(* IEC 61131-3 sources: 2026_Projet_YGO_ExcavatriceDragage/CODE_BACKUP/CODE_20260904_AvantWeekendBackup_v0.6.34/G_CYCLE (part 2) *)

(* ---- FB_CycleSemiAuto.st ---- *)
(* =======================================================================
   ⚙️ FB_CycleSemiAuto — Séquenceur du cycle automatique (Grafcet de dragage)
   ───────────────────────────────────────────────────────────────
   🎯 Rôle : Automate de cycle automatique de dragage (X0 à X13 + AX_STAB)
   🔒 Sécurité : Gating par mode et homme-mort, repli AX_STAB sur défaut
   🔌 Interface : Demandes de mouvements (treuils, translation, benne)
   📄 Doc métier : DOC/AF/AF_Partie-04_Mode_SemiAuto_Sequenceur_v2.3.md
   ======================================================================= *)

FUNCTION_BLOCK PUBLIC FB_CycleSemiAuto
VAR_INPUT
    // === COMMANDES & AUTORISATIONS ===
    Enable                  : BOOL;         // --> [CMD] Activation generale du sequenceur
    Reset                   : BOOL;         // --> [CMD] Acquittement defaut (front)
    PowerContactorEngaged   : BOOL;         // --> [SAFE] Chaine de securite OK
    EncoderFaultPresent     : BOOL;         // --> [SAFE] Defaut codeur agrege (cycle non autorise)
    Mode                    : E_Mode;       // --> [CMD] Mode arbitre (SEMI_AUTO pour instance cycle)
    JoystickDeflected       : BOOL;         // --> [CMD] Manche deflecte (non centre)
    DeadmanArmed            : BOOL;         // --> [CMD] Appui homme-mort (fenetre 3 s)
    HeartbeatIhmOk          : BOOL;         // --> [SAFE] IHM<->PLC valide

    // === COMMANDES OPERATEUR ===
    StartCycle              : BOOL;         // --> [CMD] Demande lancement / reprise (IHM)
    AbortCycle              : BOOL;         // --> [CMD] Demande abandon (IHM)

    // === CIBLES ET CONFIGURATION ===
    SelTarget               : INT;          // --> [CFG] RESERVE (C3.1 : le cycle part toujours de P1, plus de selection de cible). Cable, non consomme.
    SetDepthM               : REAL;         // --> [CFG] Profondeur de consigne (negative)
    SetOffsetM              : REAL;         // --> [CFG] Ecart de fermeture benne cible

    // === FEEDBACKS CAPTEURS & MATERIEL ===
    KoboldContactFond       : BOOL;         // --> [HW] Retour dedie Kobold : TRUE = contact fond (front descendant DI)
    KoboldImmersed          : BOOL;         // --> [HW] Etat brut DI Kobold : TRUE = sonde dans l'eau (fronts AX6/AX7)
    KoboldContactorFeedback : BOOL;         // --> [HW] Retour contacteur Kobold enclenche (verif init AX5)
    LimitLegalReached       : BOOL;         // --> [SAFE] Limite legale atteinte (descente interdite)
    LimitLegalDepthM        : REAL;         // --> [CFG] Profondeur legale minimale autorisee
    WinchSyncError          : BOOL;         // --> [SAFE] Desynchronisme bloquant M1/M2
    WinchSyncDeltaM         : REAL;         // --> [HW] Ecart codeurs M1/M2 pour diagnostic
    M1_CablePosM            : REAL;         // --> [HW] Position cable treuil M1 (recalee)
    M2_CablePosM            : REAL;         // --> [HW] Position cable treuil M2 (recalee)
    M1_MeasuredSpeedMps     : REAL;         // --> [HW] Vitesse lineaire mesuree M1 (m/s)
    M2_MeasuredSpeedMps     : REAL;         // --> [HW] Vitesse lineaire mesuree M2 (m/s)
    SpeedMismatchThresholdMps : REAL;       // --> [CFG] Seuil ecart vitesse ; 0 = controle desactive
    SpeedMismatchTimeout    : TIME;         // --> [CFG] Duree de confirmation ; 0 = controle desactive
    CableLimitM1AscentM     : REAL;         // --> [CFG] Limite haute d'exploitation M1

    // === FEEDBACKS TRANSLATION M3 ===
    Translation_At_P1           : BOOL;     // --> [HW] Capteur position P1 (arret travail)
    Translation_At_Tremie       : BOOL;     // --> [HW] Capteur fin de course tremie
    Translation_At_Maintenance : BOOL;     // --> [HW] Capteur fin de course maintenance
    Translation_Busy            : BOOL;     // --> [HW] Mouvement translation en cours
    Translation_Done            : BOOL;     // --> [HW] Cible translation atteinte

    // === FEEDBACKS BENNE ===
    Benne_Busy              : BOOL;         // --> [HW] Mouvement machoires benne en cours
    Benne_Done              : BOOL;         // --> [HW] Mouvement ouverture/fermeture termine
    Benne_IsOpen            : BOOL;         // --> [HW] Benne mecaniquement ouverte memorisee
    Benne_IsClosed          : BOOL;         // --> [HW] Benne mecaniquement fermee memorisee
    Benne_IsRoughlyClosed   : BOOL;         // --> [HW] Benne a peu pres fermee (tolerance matiere)

    // === REFERENCEMENT CODEURS ===
    HomedM1                 : BOOL;         // --> [HW] Codeur M1 reference
    HomedM2                 : BOOL;         // --> [HW] Codeur M2 reference
    TopPositionSensor       : BOOL;         // --> [HW] Capteur position haute (referencement)
    HomingRequest           : BOOL;         // --> [CMD] Demande de referencement (front)
    InitPositionOk          : BOOL;         // --> [HW] Posture de depart OK (treuils/M3 dans la plage, calcul PRG_03) - condition AX1_INIT
    WinchesAtTopWindow      : BOOL;         // --> [HW] Treuils M1 ET M2 dans la fenetre FDC logiciel haut (calcul PRG_03) - surveille en AX2

    // === CONFIG & COMMANDES CYCLE (IHM) ===
    CfgDrainTime           : TIME;         // --> [CFG] Duree d'egouttage AX13 configurable IHM (<= 0 -> defaut interne)
    SkipDrainRequest       : BOOL;         // --> [CMD] Bouton IHM : passer l'etape d'egouttage AX13 (front)
    RepositionRequest      : BOOL;         // --> [CMD] Option IHM (maintenue) : repositionnement couple M1+M2 pendant le vidage tremie (AX15B <-> AX15C)

    // === CONFIG DIVING / EXTRACTION (GEL 2026-09-03) ===
    DiveStartMinM          : REAL;         // --> [CFG] Altimetrie de lancement Kobold (AT4 : AX4 -> AX5), reglable IHM (~3..5 m ; <= 0 -> defaut interne)
    CfgRaiseOffBottomM     : REAL;         // --> [CFG] Decollement du fond en AX8 : RaiseTargetM = TouchPositionM + ce champ (reglable IHM ; <= 0 -> 0,5 m)
    CfgCtrlAscentMaxStep   : INT;          // --> [CFG] Palier max montee controle AX11, borne [1..2] (defaut 1)
    M1_SpeedStepApplied    : INT;          // --> [HW] Palier vitesse effectivement applique M1 (0 = inconnu ; garde palier <> 4 en diving)
    M2_SpeedStepApplied    : INT;          // --> [HW] Palier vitesse effectivement applique M2 (0 = inconnu)
END_VAR
VAR_OUTPUT
    // === ETATS IEC & DEFECTUOSITES ===
    Ready                   : BOOL;         // <-- [STAT] Sequenceur disponible
    Fault                   : ST_Fault;     // <-- [SAFE] Socle defaut transverse (live + latche)
    Lifecycle               : ST_Lifecycle; // <-- [STAT] Cycle de vie (Busy, Done, Waiting)
    SpeedMismatchMps        : REAL;         // <-- [DIAG] Ecart absolu vitesse M1/M2 (m/s)
    SpeedMismatchActive     : BOOL;         // <-- [DIAG] Seuil vitesse depasse sur cycle courant
    SpeedMismatchConfirmed  : BOOL;         // <-- [DIAG] Ecart vitesse confirme pendant timeout
    BottomTouched           : BOOL;         // <-- [STAT] Fond touche (latch AX8, efface a AX0 / AX_STAB / Reset) - variable d'info GEL AX8

    // === ORDRES ACTIONNEURS (COMMANDES STRUCTUREES) ===
    // Types de contrat inter-PRG uniques (ST_Program*Request) : FB_CycleSemiAuto produit
    // directement les demandes consommées par PRG_04/05/07 — plus de DUT
    // ST_fbCycle_*CmdDemand redondants ni de re-mapping champ-à-champ (NC-090).
    WinchM1Cmd              : ST_ProgramWinchRequest;        // <-- [ACT] Demande treuil M1
    WinchM2Cmd              : ST_ProgramWinchRequest;        // <-- [ACT] Demande treuil M2
    TranslationCmd          : ST_ProgramTranslationRequest;  // <-- [ACT] Demande translation M3
    BucketCmd               : ST_ProgramBucketRequest;       // <-- [ACT] Demande benne

    // === METADONNEES & SYNOPTIQUE ===
    CycleStep               : E_AutoCycleStep;          // <-- [STAT] Etape active du Grafcet
    CycleStateStr           : STRING(80);           // <-- [STAT] Libelle en clair de l'etape
    CycleStepAtError        : E_AutoCycleStep;          // <-- [DIAG] Etape specifique au moment du defaut
    OperatorActionId        : WORD;                 // <-- [DIAG] ID action operateur requise
    OperatorAction          : STRING(120);          // <-- [DIAG] Message explicatif pour l'IHM
    ExpectedAxis            : E_OperatorAxis;       // <-- [STAT] Organe joystick/bouton attendu
    ExpectedDirection       : INT;                  // <-- [STAT] Sens attendu (-1, 0, +1)
    WaitingForOperator      : BOOL;                 // <-- [STAT] En attente d'une action operateur
    WaitingForProcess       : BOOL;                 // <-- [STAT] En attente d'une condition procede
    RequestActive           : BOOL;                 // <-- [STAT] Demande de mouvement active
    CurrentCycleElapsed     : TIME;                 // <-- [DIAG] Duree ecoulee du cycle en cours (chronometre sur Lifecycle.Busy)
    LastCycleDuration       : TIME;                 // <-- [DIAG] Duree du dernier cycle acheve (figee a X13, persiste au cycle suivant)
END_VAR
VAR_IN_OUT
    // === STRUCTURES PARTAGEES & COMPTEURS ===
    SampleCount             : INT;          // <-> [BUS] Compteur de prelevements (RETAIN)
END_VAR
VAR
    // === DETECTEURS DE FRONTS ===
    ResetEdge               : R_TRIG;       // . [LOC] Detecteur front montant Reset
    StartEdge               : R_TRIG;       // . [LOC] Detecteur front montant StartCycle
    DeadmanArmedEdge        : R_TRIG;       // . [LOC] Detecteur front montant DeadmanArmed (demarrage joystick)
    AbortEdge               : R_TRIG;       // . [LOC] Detecteur front montant AbortCycle
    ErrorEdge               : R_TRIG;       // . [LOC] Detecteur front montant Error
    JoyDeflectedEdge        : R_TRIG;       // . [LOC] Front montant JoystickDeflected (relance AX18 sur geste franc, pas maintien)

    // === GATE CONTINU HOMME-MORT ===
    CycleMotionPermit       : BOOL; // . [LOC] Permis de mouvement cycle = JoystickDeflected AND DeadmanArmed (manche deflechi + homme-mort arme) ; gate commun a toutes les commandes d'actionneur du sequenceur. Le sens du mouvement reste porte par ReqAscent/ReqDescend de chaque etape.

    // === COMPTEUR PRELEVEMENTS (garde de front) ===
    SampleCountDone         : BOOL := FALSE; // . [LOC] F2: front de comptage SampleCount (1 seul increment par cycle)

    // === ETATS INTERNES ===
    State                   : E_AutoCycleStep := E_AutoCycleStep.AX0_REPOS; // . [LOC] Etape courante machine d'etat
    SavedState              : E_AutoCycleStep := E_AutoCycleStep.AX0_REPOS; // . [LOC] Etape memorisee
    PausedState             : E_AutoCycleStep := E_AutoCycleStep.AX0_REPOS; // . [LOC] Etape en pause lors de la bascule hors auto
    WaitingResume           : BOOL := FALSE;                             // . [LOC] En attente de validation consciente pour reprendre

    // === MEMORISATIONS & REGISTRES INTERNES ===
    TouchPositionM          : REAL;         // . [LOC] Position M1 memorisee lors du contact fond
    RaiseTargetM            : REAL;         // . [LOC] Profondeur de remontee memorisee
    SelectedWorkTarget      : INT;          // . [LOC] Cible de travail (fige a 3=P1 depuis C3.1) - conserve pour diag/futur
    InitConditionsOk        : BOOL;         // . [LOC] AX1_INIT : toutes les conditions initiales sont remplies
    StepMaxPrevState        : E_AutoCycleStep;  // . [LOC] Etape du scan precedent (rearmement StepMaxTimer au changement d'etape)

    // === FRONTS / TEMPO DIVING ===
    KoboldRiseEdge          : R_TRIG;       // . [LOC] Front DI Kobold 0->1 (entree dans l'eau, AX6)
    KoboldFallEdge          : F_TRIG;       // . [LOC] Front DI Kobold 1->0 (fond, AX7)
    KoboldInitTimer         : TON;          // . [LOC] Fenetre de verif retour contacteur Kobold en AX5
    RetryJoyReleaseTimer    : TON;          // . [LOC] Anti-rebond relache joystick pendant diving (>= 200 ms avant reprise)
    PalierNot4Timer         : TON;          // . [LOC] Confirmation palier bloque < 4 en plongee (tolere la rampe 1->4)
    DivingRetryTrig         : BOOL;         // . [LOC] Synthese GT-dive-retry (erreur Kobold / joystick relache / palier < 4 confirme en AX5..AX7)
    CtrlAscentMaxStepEff    : INT;          // . [LOC] CfgCtrlAscentMaxStep borne [1..2]
    RaiseOffBottomEff       : REAL;         // . [LOC] CfgRaiseOffBottomM borne (>0, defaut 0,5 m)
    DiveStartMinEff         : REAL;         // . [LOC] DiveStartMinM borne (defaut interne si <= 0)

    // === TEMPORISATEURS INTERNES ===
    DrainingTimer           : TON;          // . [LOC] Temporisateur de vidage (egouttage), PT = DrainTimeEff
    CycleRunTimer           : TON;          // . [LOC] Chronometre du cycle en cours (IN = Lifecycle.Busy) ; .ET = duree
    SkipDrainEdge           : R_TRIG;       // . [LOC] Front bouton IHM "passer egouttage"
    DrainTimeEff            : TIME;         // . [LOC] Duree d'egouttage effective (CfgDrainTime bornee au defaut interne)
    StabilizationTimer      : TON;          // . [LOC] Temporisation maximale de remontee lente
    SpeedMismatchTimer      : TON;          // . [LOC] Confirmation temporelle ecart de vitesse
    StepMaxTimer            : TON;          // . [LOC] Tempo max d'etape

    // === CONSTANTES & CONFIGURATIONS INTERNES ===
    CtrlAscentDistM         : REAL := 2.0;      // . [LOC] Distance de remontee lente de controle
    CtrlAscentToleranceM    : REAL := 0.25;     // . [LOC] Ecart maximal admis entre codeurs
    CtrlAscentTimeout       : TIME := T#30s;    // . [LOC] Temps max pour zone de stabilisation
    DrainingTime            : TIME := T#5s;     // . [LOC] Temps d'egouttage par defaut
    StepMaxTimeout          : TIME := T#60s;    // . [LOC] Tempo max d'etape

    // === SOCLE DEFAUT TRANSVERSE ===
    instFault               : FB_FaultCore;                  // * [INST] Socle defaut transverse
    instCauses              : ARRAY[0..15] OF ST_FaultCause; // . [LOC] Table des causes de defaut
END_VAR
VAR CONSTANT
    // Paliers de vitesse treuil par etape (StepTgt des demandes WinchMxCmd, 1..5 ; 0 = arret).
    CST_StepSlow   : INT := 1;   // Palier lent : retente AX9, controle AX11, repositionnement AX15C
    CST_StepDive   : INT := 4;   // Palier plongee Kobold AX4..AX7 : palier 4 MINI ET MAXI impose, palier 5 interdit (GEL Q9)
    CST_StepLoaded : INT := 4;   // Palier montee en charge AX12 (bridage strict <= 4, jamais palier 5)
    CST_KoboldInitTimeout : TIME := T#3s;   // Fenetre max de confirmation retour contacteur Kobold en AX5
    CST_RaiseOffBottomDefaultM : REAL := 0.5;   // Decollement du fond par defaut (AX8) si CfgRaiseOffBottomM <= 0
    // Backstop anti-telescopage : ecart de position M1/M2 max tolere pendant les phases
    // reellement couplees hors X7 (qui a deja son propre controle a 0,25 m). Aligne sur
    // CfgSyncCriticalToleranceM = 0,50 m (AF-04 §5). FB_SyncDeviation (PRG_04) reste la
    // surveillance primaire ; ceci est un garde-fou local au sequenceur.
    CST_CoupledPosBacklashM : REAL := 0.5;
END_VAR

// === IMPLEMENTATION ===

{region "§1 Causes & Socle Défaut"}
// 🔑 1. FRONTS ET CAUSES
ResetEdge(CLK := Reset);
StartEdge(CLK := StartCycle);
DeadmanArmedEdge(CLK := DeadmanArmed);
AbortEdge(CLK := AbortCycle);
SkipDrainEdge(CLK := SkipDrainRequest);
KoboldRiseEdge(CLK := KoboldImmersed);
KoboldFallEdge(CLK := KoboldImmersed);
JoyDeflectedEdge(CLK := JoystickDeflected);

// Config diving/extraction bornee (repli defaut interne si non reglee / valeur implausible).
// DiveStartMinM = altimetrie de lancement Kobold dans le referentiel M1_CablePosM
// (positif, ~7,5 m au FDC haut, decroissant a la descente). Plage plausible 0,5..8,0 m ;
// hors plage -> repli 4,0 m.
IF (DiveStartMinM >= 0.5) AND (DiveStartMinM <= 8.0) THEN
    DiveStartMinEff := DiveStartMinM;
ELSE
    DiveStartMinEff := 4.0;
END_IF;
RaiseOffBottomEff := SEL(CfgRaiseOffBottomM > 0.0, CST_RaiseOffBottomDefaultM, CfgRaiseOffBottomM);
CtrlAscentMaxStepEff := LIMIT(1, CfgCtrlAscentMaxStep, 2);

// ⏱️ Chronomètre du cycle : compte tant que le séquenceur est actif (Lifecycle.Busy).
// .ET = durée écoulée du cycle en cours ; figée dans LastCycleDuration à l'achèvement (X13).
CycleRunTimer(IN := Lifecycle.Busy, PT := T#12h);
CurrentCycleElapsed := CycleRunTimer.ET;

// Durée d'égouttage effective : config IHM si valide, sinon défaut interne.
DrainTimeEff := SEL(CfgDrainTime <= T#0s, CfgDrainTime, DrainingTime);

// ⏱️ Surveillance indépendante de la remontée lente de controle
// AX11_CTRL_ASCENT -> AX12_LOADED_ASCENT : TON de stabilisation palier lent.
StabilizationTimer(IN := (State = E_AutoCycleStep.AX11_CTRL_ASCENT), PT := CtrlAscentTimeout);

// ⏱️ AX5_KOBOLD_INIT : fenetre de confirmation du retour contacteur Kobold.
KoboldInitTimer(IN := (State = E_AutoCycleStep.AX5_KOBOLD_INIT), PT := CST_KoboldInitTimeout);

// 📏 Comparaison vitesse réelle M1/M2
SpeedMismatchMps := ABS(M1_MeasuredSpeedMps - M2_MeasuredSpeedMps);
SpeedMismatchActive := (State = E_AutoCycleStep.AX11_CTRL_ASCENT)
                       AND JoystickDeflected
                       AND (SpeedMismatchThresholdMps > 0.0)
                       AND (SpeedMismatchTimeout > T#0ms)
                       AND (SpeedMismatchMps > SpeedMismatchThresholdMps);
// AX11_CTRL_ASCENT -> AX_STAB : TON confirmation écart vitesse.
SpeedMismatchTimer(IN := SpeedMismatchActive, PT := SpeedMismatchTimeout);
SpeedMismatchConfirmed := SpeedMismatchTimer.Q;

// Tempo max d'étape (R5) — backstop durée d'état, lancé SEULEMENT si pilotage joystick actif.
// Xi -> AX_STAB sur dépassement. Réarmé à CHAQUE changement d'étape (IN=FALSE 1 scan) :
// chaque étape dispose de sa propre fenêtre StepMaxTimeout, la tempo n'est PAS cumulative
// sur l'ensemble du cycle (un cycle réel long ne tombe plus en AX_STAB intempestif).
StepMaxTimer(IN := (State = StepMaxPrevState)
                  AND JoystickDeflected
                  AND (State <> E_AutoCycleStep.AX0_REPOS)
                  AND (State <> E_AutoCycleStep.AX18_DONE_SYNC)
                  AND (State <> E_AutoCycleStep.AX_STAB)
                  AND (State <> E_AutoCycleStep.AX_DIVING_RETRY),
             PT := StepMaxTimeout);
StepMaxPrevState := State;

// Egouttage AX13 : TON gaté sur l'étape (remis à 0 hors AX13). Remplace l'ancien IN:=TRUE câblé
// qui pouvait laisser Q déjà vrai à l'entrée en AX13 (temps d'égouttage non respecté).
DrainingTimer(IN := (State = E_AutoCycleStep.AX13_DRAIN_PAUSE), PT := DrainTimeEff);

// GT-dive-retry (GEL Q11) : en AX5/AX6/AX7, erreur sequence Kobold (retour contacteur
// absent apres CST_KoboldInitTimeout) OU joystick relache (>= 200 ms, anti-rebond) OU
// palier applique <> 4 sur M1 ou M2 (feedback si cable) -> reprise AX_DIVING_RETRY
// (PAS un defaut latche).
RetryJoyReleaseTimer(IN := ((State = E_AutoCycleStep.AX5_KOBOLD_INIT)
                             OR (State = E_AutoCycleStep.AX6_SEARCH_IMMERSION)
                             OR (State = E_AutoCycleStep.AX7_SEARCH_BOTTOM))
                            AND NOT JoystickDeflected,
                     PT := T#200ms);
// Palier bloque SOUS 4 pendant la plongee : on TOLERE la rampe 1->4 (tempo contacteurs,
// GEL AX4) ; seul un blocage confirme > 4 s en AX5..AX7 declenche la reprise. Palier 5
// (> 4) est traite instantanement par la cause de defaut 8 (latche), pas ici.
PalierNot4Timer(IN := ((State = E_AutoCycleStep.AX5_KOBOLD_INIT)
                        OR (State = E_AutoCycleStep.AX6_SEARCH_IMMERSION)
                        OR (State = E_AutoCycleStep.AX7_SEARCH_BOTTOM))
                       AND JoystickDeflected
                       AND ( ((M1_SpeedStepApplied > 0) AND (M1_SpeedStepApplied < CST_StepDive))
                          OR ((M2_SpeedStepApplied > 0) AND (M2_SpeedStepApplied < CST_StepDive)) ),
                PT := T#5s);
DivingRetryTrig := ((State = E_AutoCycleStep.AX5_KOBOLD_INIT)
                     OR (State = E_AutoCycleStep.AX6_SEARCH_IMMERSION)
                     OR (State = E_AutoCycleStep.AX7_SEARCH_BOTTOM))
                   AND ( (KoboldInitTimer.Q AND NOT KoboldContactorFeedback)
                         OR RetryJoyReleaseTimer.Q
                         OR PalierNot4Timer.Q );

// Table des causes de défaut
instCauses[0].Active   := LimitLegalReached
                          AND ((State = E_AutoCycleStep.AX4_DESCEND_DIVING)
                            OR (State = E_AutoCycleStep.AX5_KOBOLD_INIT)
                            OR (State = E_AutoCycleStep.AX6_SEARCH_IMMERSION)
                            OR (State = E_AutoCycleStep.AX7_SEARCH_BOTTOM));
instCauses[0].Latching := TRUE;
instCauses[0].Texte    := 'Limite legale de profondeur atteinte pendant descente';

instCauses[1].Active   := WinchSyncError AND (State <> E_AutoCycleStep.AX0_REPOS) AND (State <> E_AutoCycleStep.AX_STAB);
instCauses[1].Latching := TRUE;
instCauses[1].Texte    := 'Desynchronisme treuils M1/M2 bloquant';

instCauses[2].Active   := SpeedMismatchConfirmed AND (State <> E_AutoCycleStep.AX0_REPOS) AND (State <> E_AutoCycleStep.AX_STAB);
instCauses[2].Latching := TRUE;
instCauses[2].Texte    := 'Ecart de vitesse M1/M2 confirme en montee';

instCauses[3].Active   := NOT HeartbeatIhmOk AND (State <> E_AutoCycleStep.AX0_REPOS) AND (State <> E_AutoCycleStep.AX_STAB);
instCauses[3].Latching := TRUE;
instCauses[3].Texte    := 'Perte communication IHM pendant cycle';

instCauses[4].Active   := StepMaxTimer.Q AND (State <> E_AutoCycleStep.AX_STAB);
instCauses[4].Latching := TRUE;
instCauses[4].Texte    := 'Depassement tempo maximale d etape (blocage mouvement)';

instCauses[5].Active   := (StabilizationTimer.Q OR (ABS(M1_CablePosM - M2_CablePosM) > CtrlAscentToleranceM))
                          AND (State = E_AutoCycleStep.AX11_CTRL_ASCENT);
instCauses[5].Latching := TRUE;
instCauses[5].Texte    := 'Defaut de stabilisation / tolerance ecart codeurs en remontee controle';

// Backstop anti-telescopage : ecart de position M1/M2 excessif pendant une phase
// reellement couplee. AX11 a deja son propre controle (instCauses[5]). Seuil grossier
// (0,50 m) : filet local si FB_SyncDeviation (PRG_04) ne coupe pas.
instCauses[6].Active   := (ABS(M1_CablePosM - M2_CablePosM) > CST_CoupledPosBacklashM)
                          AND JoystickDeflected
                          AND ((State = E_AutoCycleStep.AX4_DESCEND_DIVING)
                            OR (State = E_AutoCycleStep.AX5_KOBOLD_INIT)
                            OR (State = E_AutoCycleStep.AX6_SEARCH_IMMERSION)
                            OR (State = E_AutoCycleStep.AX7_SEARCH_BOTTOM)
                            OR (State = E_AutoCycleStep.AX9_RAISE_OFF_BOTTOM)
                            OR (State = E_AutoCycleStep.AX12_LOADED_ASCENT)
                            OR (State = E_AutoCycleStep.AX15C_DUMP_REPOSITION));
instCauses[6].Latching := TRUE;
instCauses[6].Texte    := 'Ecart de position M1/M2 excessif en phase couplee (anti-telescopage)';

// AX2 : pendant la translation vers P1 les treuils M1/M2 doivent RESTER au FDC
// logiciel haut (WinchesAtTopWindow, calcul PRG_03). S'ils quittent la fenetre
// -> defaut latche, sortie cycle (GEL SEMI_AUTO cause 7 / Q10).
instCauses[7].Active   := NOT WinchesAtTopWindow AND (State = E_AutoCycleStep.AX2_TRANSLATE_P1);
instCauses[7].Latching := TRUE;
instCauses[7].Texte    := 'Treuils M1/M2 hors FDC haut pendant la translation vers P1';

// GEL cause 8 : palier vitesse > 4 (palier 5) applique pendant la plongee. Le FB commande
// toujours CST_StepDive = 4 ; un palier 5 en retour feedback = anomalie aval -> defaut latche.
// (Un palier < 4 en retour est traite en reprise par GT-dive-retry, pas ici.)
instCauses[8].Active   := (((M1_SpeedStepApplied > CST_StepDive) OR (M2_SpeedStepApplied > CST_StepDive)))
                          AND ((State = E_AutoCycleStep.AX4_DESCEND_DIVING)
                            OR (State = E_AutoCycleStep.AX5_KOBOLD_INIT)
                            OR (State = E_AutoCycleStep.AX6_SEARCH_IMMERSION)
                            OR (State = E_AutoCycleStep.AX7_SEARCH_BOTTOM));
instCauses[8].Latching := TRUE;
instCauses[8].Texte    := 'Palier vitesse > 4 (palier 5) pendant la plongee - interdit';

// Appel du socle de défaut
instFault(Enable := Enable, Reset := Reset, Causes := instCauses);
Fault := instFault.Fault;
ErrorEdge(CLK := Fault.Error);
{endregion}

{region "§2 Gate securite & Bascule Mode"}
// 🛑 2. GATES DE SÉCURITÉ ET NEUTRALISATION
// Le mode SEMI_AUTO peut être sélectionné sous AU/défaut (FB_Modes), mais le cycle
// ne tourne JAMAIS sans puissance (PowerContactorEngaged) ni avec un codeur défaillant
// (EncoderFaultPresent) — les données de position invalides rendraient le Grafcet erroné.
IF NOT Enable OR NOT PowerContactorEngaged OR EncoderFaultPresent THEN
    WinchM1Cmd.RunRequest     := FALSE;
    WinchM1Cmd.ReqAscent      := FALSE;
    WinchM1Cmd.ReqDescend     := FALSE;
    WinchM1Cmd.StepTgt        := 0;

    WinchM2Cmd.RunRequest     := FALSE;
    WinchM2Cmd.ReqAscent      := FALSE;
    WinchM2Cmd.ReqDescend     := FALSE;
    WinchM2Cmd.StepTgt        := 0;

    TranslationCmd.ReqStart   := FALSE;
    TranslationCmd.PositionTgt  := 0;

    BucketCmd.ReqOpen         := FALSE;
    BucketCmd.ReqClose        := FALSE;
    BucketCmd.ReqKoboldMeasureEnable := FALSE;

    // Si on quitte le semi-auto alors qu'un cycle était en cours, on mémorise l'étape pour la pause
    IF (State <> E_AutoCycleStep.AX0_REPOS) AND (State <> E_AutoCycleStep.AX18_DONE_SYNC) AND (State <> E_AutoCycleStep.AX_STAB) THEN
        PausedState := State;
        WaitingResume := TRUE;
    END_IF;

    CycleStep            := State;
    CycleStateStr        := 'Cycle desactive : securite/codeur/mode';
    Ready                := FALSE;
    Lifecycle.Busy       := FALSE;
    Lifecycle.Done       := FALSE;
    SpeedMismatchTimer(IN := FALSE, PT := SpeedMismatchTimeout);
    SpeedMismatchMps := 0.0;
    SpeedMismatchActive := FALSE;
    SpeedMismatchConfirmed := FALSE;
    OperatorActionId := 0;
    IF EncoderFaultPresent THEN
        OperatorAction := 'Cycle non autorise : defaut codeur present. Reinitialiser le defaut codeur.';
    ELSE
        OperatorAction := 'Passer en mode Semi-Auto et engager la securite pour activer le cycle.';
    END_IF;
    ExpectedAxis := E_OperatorAxis.NONE;
    ExpectedDirection := 0;
    WaitingForOperator := FALSE;
    WaitingForProcess := FALSE;
    RequestActive := FALSE;
    RETURN;
END_IF;

Ready := Enable AND NOT Fault.Latched;

// 🛡️ Gate continu homme-mort : le mouvement n'est autorisé que si le manche est
// défléchi (JoystickDeflected) ET l'homme-mort est armé (DeadmanArmed). Chaque
// commande de mouvement est gatée par ce permis à chaque scan (pas seulement au
// démarrage). Le séquenceur (transitions X0→X13) reste piloté par JoystickDeflected.
CycleMotionPermit := JoystickDeflected AND DeadmanArmed;

// Au retour en Semi-Auto, si une étape était en cours, on exige une reprise consciente
IF WaitingResume THEN
    // 🔒 Sécurité anti-redémarrage automatique (AF-04 §4.1) : le cycle ne reprend
    // PAS sur manche + homme-mort seuls. Il reste en attente d'un geste conscient
    // (StartCycle) avant de restaurer l'étape mémorisée.
    IF StartEdge.Q THEN
        State := PausedState;   // reprise consciente : restaure l'étape mémorisée
        WaitingResume := FALSE;
    ELSE
        // Hold : neutralise toute demande de mouvement et affiche l'attente.
        WinchM1Cmd.RunRequest := FALSE; WinchM1Cmd.ReqAscent := FALSE; WinchM1Cmd.ReqDescend := FALSE; WinchM1Cmd.StepTgt := 0;
        WinchM2Cmd.RunRequest := FALSE; WinchM2Cmd.ReqAscent := FALSE; WinchM2Cmd.ReqDescend := FALSE; WinchM2Cmd.StepTgt := 0;
        TranslationCmd.ReqStart := FALSE; TranslationCmd.PositionTgt := 0;
        BucketCmd.ReqOpen := FALSE; BucketCmd.ReqClose := FALSE; BucketCmd.ReqKoboldMeasureEnable := FALSE;
        CycleStep := PausedState;
        CycleStateStr := 'Cycle en pause : reprise consciente requise (StartCycle)';
        Lifecycle.Busy := FALSE;
        Lifecycle.Done := FALSE;
        ExpectedAxis := E_OperatorAxis.BUTTON;
        ExpectedDirection := 0;
        WaitingForOperator := TRUE;
        WaitingForProcess := FALSE;
        OperatorActionId := 16#0400;
        OperatorAction := 'Reprendre le cycle : appuyer sur StartCycle (geste conscient).';
        RequestActive := FALSE;
    END_IF;
END_IF;

// 🧊 R9 — capture l'étape spécifique AVANT la bascule vers AX_STAB
IF ErrorEdge.Q THEN
    CycleStepAtError := State;
    State := E_AutoCycleStep.AX_STAB;
    WaitingResume := FALSE;   // un défaut abroge la reprise consciente : repli AX_STAB
END_IF;

// GT-dive-retry (GEL Q11) : reprise de plongee (PAS un defaut latche). Prioritaire
// apres le repli defaut : une vraie erreur (ErrorEdge) l'emporte.
IF DivingRetryTrig AND (State <> E_AutoCycleStep.AX_STAB) THEN
    State := E_AutoCycleStep.AX_DIVING_RETRY;
END_IF;

IF ResetEdge.Q THEN
    SavedState := E_AutoCycleStep.AX0_REPOS;
    BottomTouched := FALSE;
    IF State = E_AutoCycleStep.AX_STAB THEN
        State := E_AutoCycleStep.AX0_REPOS;
    END_IF;
END_IF;

// Gestion de l'Abandon explicite
IF AbortEdge.Q THEN
    State := E_AutoCycleStep.AX0_REPOS;
    WaitingResume := FALSE;
    PausedState := E_AutoCycleStep.AX0_REPOS;
END_IF;

// SEMI_AUTO : FB_CycleSemiAuto est le SEUL producteur des demandes benne. Les champs
// assistants (DiveSearch/ExtractionAssist) sont inactifs en cycle automatique
// -> valeurs neutres déterministes (identiques à la branche SEMI_AUTO de PRG_03).
BucketCmd.DescendPermitDiveBucketOpen := TRUE;
BucketCmd.ExtractionControlActive := FALSE;
BucketCmd.MinStepDown := 0;
{endregion}

{region "§3 Machine etat cycle automatique"}
// 🔁 2. LOGIQUE DU SÉQUENCEUR (Machine d'état) — CASE sur enum unique (R1)
// Pendant une reprise consciente (WaitingResume), le séquenceur est gelé :
// l'étape mémorisée ne s'exécute pas tant que StartCycle n'a pas été appuyé.
IF NOT WaitingResume THEN
CASE State OF

    E_AutoCycleStep.AX0_REPOS:
        CycleStep := E_AutoCycleStep.AX0_REPOS;
        CycleStateStr := 'AX0 - Verification coherence systeme';
        WinchM1Cmd.RunRequest := FALSE; WinchM1Cmd.ReqAscent := FALSE; WinchM1Cmd.ReqDescend := FALSE; WinchM1Cmd.StepTgt := 0;
        WinchM2Cmd.RunRequest := FALSE; WinchM2Cmd.ReqAscent := FALSE; WinchM2Cmd.ReqDescend := FALSE; WinchM2Cmd.StepTgt := 0;
        TranslationCmd.ReqStart := FALSE; TranslationCmd.PositionTgt := 0;
        BucketCmd.ReqOpen := FALSE; BucketCmd.ReqClose := FALSE; BucketCmd.ReqKoboldMeasureEnable := FALSE;
        Lifecycle.Busy := FALSE;
        Lifecycle.Done := FALSE;
        ExpectedAxis := E_OperatorAxis.BUTTON;
        ExpectedDirection := 0;
        WaitingForOperator := TRUE;
        WaitingForProcess := FALSE;
        OperatorActionId := 16#0400;
        OperatorAction := 'AX0 - Demander le demarrage du cycle (Bouton IHM ou armement Homme-Mort).';
        SampleCountDone := FALSE;   // F2: réarmement du front de comptage à chaque entrée en X0
        BottomTouched   := FALSE;   // info fond touche effacee au repos

        // Transition si système sain et réarmé (front reset ou démarrage).
        // 🔫 D2 : démarrage par bouton IHM (StartEdge) OU armement homme-mort joystick
        IF (StartEdge.Q OR DeadmanArmedEdge.Q) AND NOT Fault.Latched THEN
            WaitingResume := FALSE;
            State := E_AutoCycleStep.AX1_INIT;
        END_IF;

    E_AutoCycleStep.AX1_INIT:
        CycleStep := E_AutoCycleStep.AX1_INIT;
        Lifecycle.Busy := TRUE;
        Lifecycle.Done := FALSE;
        ExpectedDirection := 0;

        // AX1_INIT : verification des CONDITIONS INITIALES du cycle. AUCUN ordre de
        // mouvement, aucun referencement (datum M1/M2/benne = responsabilite exclusive
        // FB_CycleMachineHoming). Conditions : codeurs M1/M2 references, aucun defaut
        // latche, treuils au FDC logiciel haut (TopPositionSensor), et posture de depart
        // OK (InitPositionOk : chariot M3 PAS a droite de P1 + treuils dans la plage
        // +/- 0,4 m autour du FDC haut, calcul PRG_03 ; positionnement fin P1 = AX2).
        InitConditionsOk := HomedM1 AND HomedM2 AND NOT Fault.Latched
                            AND TopPositionSensor AND InitPositionOk;
        IF InitConditionsOk THEN
            CycleStateStr := 'AX1 - Conditions initiales OK';
            ExpectedAxis := E_OperatorAxis.NONE;
            WaitingForOperator := FALSE;
            WaitingForProcess := TRUE;
            OperatorActionId := 0;
            OperatorAction := '';
            State := E_AutoCycleStep.AX2_TRANSLATE_P1;   // franchie sans mouvement
        ELSIF NOT (HomedM1 AND HomedM2) THEN
            CycleStateStr := 'AX1 - Machine non referencee';
            ExpectedAxis := E_OperatorAxis.BUTTON;
            WaitingForOperator := TRUE;
            WaitingForProcess := FALSE;
            OperatorActionId := 16#0401;
            OperatorAction := 'AX1 - Machine non referencee : passer en maintenance pour le referencement.';
        ELSE
            CycleStateStr := 'AX1 - Conditions initiales non remplies';
            ExpectedAxis := E_OperatorAxis.BUTTON;
            WaitingForOperator := TRUE;
            WaitingForProcess := FALSE;
            OperatorActionId := 16#0401;
            OperatorAction := 'AX1 - Amener les treuils au FDC haut.';
        END_IF;

    E_AutoCycleStep.AX2_TRANSLATE_P1:
        CycleStep := E_AutoCycleStep.AX2_TRANSLATE_P1;
        CycleStateStr := 'AX2 - Mise en position P1 (translation)';
        Lifecycle.Busy := TRUE;
        Lifecycle.Done := FALSE;
        ExpectedAxis := E_OperatorAxis.JOYSTICK_X;
        // GEL SEMI_AUTO Q10 : le cycle n'emet AUCUNE commande M3 automatique (pas de
        // selection de cible). L'operateur pousse le joystick VERS LA DROITE et amene M3
        // a P1 ; ralenti PV + arret sur FDC P1 assures par PRG_05/FB_Translation (comme en
        // maintenance). Le cycle SURVEILLE en permanence que les treuils M1/M2 RESTENT au
        // FDC logiciel haut (WinchesAtTopWindow) : sortie sur defaut latche (cause 7) sinon.
        // Le controle "chariot pas a droite de P1" est fait en AX1_INIT, pas ici.
        WinchM1Cmd.RunRequest := FALSE; WinchM1Cmd.ReqAscent := FALSE; WinchM1Cmd.ReqDescend := FALSE; WinchM1Cmd.StepTgt := 0;
        WinchM2Cmd.RunRequest := FALSE; WinchM2Cmd.ReqAscent := FALSE; WinchM2Cmd.ReqDescend := FALSE; WinchM2Cmd.StepTgt := 0;
        TranslationCmd.PositionTgt := 3;          // repere P1 pour PRG_05 (info ; pas de pilotage cycle)

        IF Translation_At_P1 THEN
            ExpectedDirection := 0;
            WaitingForOperator := FALSE;
            WaitingForProcess := TRUE;
            OperatorActionId := 16#0402;
            OperatorAction := 'AX2 - Position P1 atteinte.';
            TranslationCmd.ReqStart := FALSE;
            State := E_AutoCycleStep.AX3_OPEN_BUCKET;
        ELSE
            // Entre tremie et P1 : l'operateur pousse le joystick VERS LA DROITE (axe
            // Tremie--P2--P1--Maintenance : P1 est a droite de la tremie). Maintien requis ;
            // ralenti PV + arret FDC P1 assures par PRG_05. Transition sur P1 STABILISE.
            ExpectedDirection := 1;
            WaitingForOperator := NOT JoystickDeflected;
            WaitingForProcess := JoystickDeflected;
            OperatorActionId := 16#0402;
            OperatorAction := 'AX2 - Pousser le joystick vers la droite : arret automatique sur P1.';
            TranslationCmd.ReqStart := CycleMotionPermit;
        END_IF;

    E_AutoCycleStep.AX3_OPEN_BUCKET:
        CycleStep := E_AutoCycleStep.AX3_OPEN_BUCKET;
        CycleStateStr := 'AX3 - Ouverture benne';
        Lifecycle.Busy := TRUE;
        Lifecycle.Done := FALSE;
        ExpectedAxis := E_OperatorAxis.JOYSTICK_Y;
        ExpectedDirection := 0;
        WaitingForOperator := NOT JoystickDeflected;
        WaitingForProcess := JoystickDeflected;
        OperatorActionId := 16#0403;
        OperatorAction := 'AX3 - Joystick pousse : ouverture benne jusqu au FDC logiciel benne ouverte.';

        // X3 = etape benne seule : treuils explicitement neutralises (config treuil unique par etape).
        WinchM1Cmd.RunRequest := FALSE; WinchM1Cmd.ReqAscent := FALSE; WinchM1Cmd.ReqDescend := FALSE; WinchM1Cmd.StepTgt := 0;
        WinchM2Cmd.RunRequest := FALSE; WinchM2Cmd.ReqAscent := FALSE; WinchM2Cmd.ReqDescend := FALSE; WinchM2Cmd.StepTgt := 0;

        IF Benne_IsOpen THEN
            State := E_AutoCycleStep.AX4_DESCEND_DIVING;
        ELSE
            BucketCmd.ReqOpen := CycleMotionPermit;
            IF JoystickDeflected AND Benne_Done AND Benne_IsOpen THEN
                BucketCmd.ReqOpen := FALSE;
                State := E_AutoCycleStep.AX4_DESCEND_DIVING;
            END_IF;
        END_IF;

    (* ===================== DIVING (AX4..AX8 + AX_DIVING_RETRY) ===================== *)

    E_AutoCycleStep.AX4_DESCEND_DIVING:
        CycleStep := E_AutoCycleStep.AX4_DESCEND_DIVING;
        CycleStateStr := 'AX4 - Plongee couplee palier 4 jusqu a l altimetrie de lancement';
        Lifecycle.Busy := TRUE;
        Lifecycle.Done := FALSE;
        ExpectedAxis := E_OperatorAxis.JOYSTICK_Y;
        ExpectedDirection := -1;
        WaitingForOperator := NOT JoystickDeflected;
        WaitingForProcess := JoystickDeflected;
        OperatorActionId := 16#0404;
        OperatorAction := 'AX4 - Maintenir la descente palier 4 (Kobold pas encore enclenche).';

        // Palier 4 MINI ET MAXI (CST_StepDive), palier 5 interdit (cause 8). Tempo
        // sequencement contacteurs conservee en aval (PRG_04 : montee progressive 1->4).
        // Contacteur Kobold PAS enclenche a cette etape.
        WinchM1Cmd.RunRequest := CycleMotionPermit;
        WinchM1Cmd.ReqAscent := FALSE; WinchM1Cmd.ReqDescend := TRUE;
        WinchM1Cmd.StepTgt  := CST_StepDive;
        WinchM2Cmd.RunRequest := CycleMotionPermit;
        WinchM2Cmd.ReqAscent := FALSE; WinchM2Cmd.ReqDescend := TRUE;
        WinchM2Cmd.StepTgt  := CST_StepDive;
        BucketCmd.ReqKoboldMeasureEnable := FALSE;

        // AT4 : altimetrie de lancement atteinte (M1 ET M2 <= DiveStartMinEff).
        IF JoystickDeflected
           AND (M1_CablePosM <= DiveStartMinEff) AND (M2_CablePosM <= DiveStartMinEff) THEN
            State := E_AutoCycleStep.AX5_KOBOLD_INIT;
        END_IF;

    E_AutoCycleStep.AX5_KOBOLD_INIT:
        CycleStep := E_AutoCycleStep.AX5_KOBOLD_INIT;
        CycleStateStr := 'AX5 - Activation contacteur Kobold au vol';
        Lifecycle.Busy := TRUE;
        Lifecycle.Done := FALSE;
        ExpectedAxis := E_OperatorAxis.JOYSTICK_Y;
        ExpectedDirection := -1;
        WaitingForOperator := NOT JoystickDeflected;
        WaitingForProcess := JoystickDeflected;
        OperatorActionId := 16#0405;
        OperatorAction := 'AX5 - Maintenir la descente palier 4 : initialisation Kobold en cours.';

        // Descente palier 4 maintenue ; enclenche le contacteur Kobold et attend le retour.
        WinchM1Cmd.RunRequest := CycleMotionPermit;
        WinchM1Cmd.ReqAscent := FALSE; WinchM1Cmd.ReqDescend := TRUE;
        WinchM1Cmd.StepTgt  := CST_StepDive;
        WinchM2Cmd.RunRequest := CycleMotionPermit;
        WinchM2Cmd.ReqAscent := FALSE; WinchM2Cmd.ReqDescend := TRUE;
        WinchM2Cmd.StepTgt  := CST_StepDive;
        BucketCmd.ReqKoboldMeasureEnable := CycleMotionPermit;

        // AT5 : retour contacteur Kobold coherent -> recherche immersion.
        // (echec init / joystick relache / palier <> 4 -> AX_DIVING_RETRY via GT-dive-retry §1)
        IF JoystickDeflected AND KoboldContactorFeedback THEN
            State := E_AutoCycleStep.AX6_SEARCH_IMMERSION;
        END_IF;

    E_AutoCycleStep.AX6_SEARCH_IMMERSION:
        CycleStep := E_AutoCycleStep.AX6_SEARCH_IMMERSION;
        CycleStateStr := 'AX6 - Recherche entree dans l eau (front DI Kobold 0->1)';
        Lifecycle.Busy := TRUE;
        Lifecycle.Done := FALSE;
        ExpectedAxis := E_OperatorAxis.JOYSTICK_Y;
        ExpectedDirection := -1;
        WaitingForOperator := NOT JoystickDeflected;
        WaitingForProcess := JoystickDeflected;
        OperatorActionId := 16#0406;
        OperatorAction := 'AX6 - Maintenir la descente palier 4 : entree dans l eau attendue.';

        WinchM1Cmd.RunRequest := CycleMotionPermit;
        WinchM1Cmd.ReqAscent := FALSE; WinchM1Cmd.ReqDescend := TRUE;
        WinchM1Cmd.StepTgt  := CST_StepDive;
        WinchM2Cmd.RunRequest := CycleMotionPermit;
        WinchM2Cmd.ReqAscent := FALSE; WinchM2Cmd.ReqDescend := TRUE;
        WinchM2Cmd.StepTgt  := CST_StepDive;
        BucketCmd.ReqKoboldMeasureEnable := CycleMotionPermit;

        // AT6 : front montant DI Kobold (immersion confirmee) -> recherche du fond.
        IF JoystickDeflected AND KoboldRiseEdge.Q THEN
            State := E_AutoCycleStep.AX7_SEARCH_BOTTOM;
        END_IF;

    E_AutoCycleStep.AX7_SEARCH_BOTTOM:
        CycleStep := E_AutoCycleStep.AX7_SEARCH_BOTTOM;
        CycleStateStr := 'AX7 - Recherche du fond (front DI Kobold 1->0)';
        Lifecycle.Busy := TRUE;
        Lifecycle.Done := FALSE;
        ExpectedAxis := E_OperatorAxis.JOYSTICK_Y;
        ExpectedDirection := -1;
        WaitingForOperator := NOT JoystickDeflected;
        WaitingForProcess := JoystickDeflected;
        OperatorActionId := 16#0407;
        OperatorAction := 'AX7 - Maintenir la descente palier 4 sous l eau : detection du fond.';

        WinchM1Cmd.RunRequest := CycleMotionPermit;
        WinchM1Cmd.ReqAscent := FALSE; WinchM1Cmd.ReqDescend := TRUE;
        WinchM1Cmd.StepTgt  := CST_StepDive;
        WinchM2Cmd.RunRequest := CycleMotionPermit;
        WinchM2Cmd.ReqAscent := FALSE; WinchM2Cmd.ReqDescend := TRUE;
        WinchM2Cmd.StepTgt  := CST_StepDive;
        BucketCmd.ReqKoboldMeasureEnable := CycleMotionPermit;

        // AT7 : front descendant DI Kobold (ou retour dedie KoboldContactFond) = fond.
        IF JoystickDeflected AND (KoboldFallEdge.Q OR KoboldContactFond) THEN
            State := E_AutoCycleStep.AX8_BOTTOM_CONFIRMED;
        END_IF;

    E_AutoCycleStep.AX8_BOTTOM_CONFIRMED:
        CycleStep := E_AutoCycleStep.AX8_BOTTOM_CONFIRMED;
        CycleStateStr := 'AX8 - Fond confirme : coupure treuils, memorisation';
        Lifecycle.Busy := TRUE;
        Lifecycle.Done := FALSE;
        ExpectedAxis := E_OperatorAxis.NONE;
        ExpectedDirection := 0;
        WaitingForOperator := FALSE;
        WaitingForProcess := TRUE;
        OperatorActionId := 16#0408;
        OperatorAction := 'AX8 - Fond touche.';

        // Coupure INSTANTANEE de toutes les commandes treuils (meme scan) + Kobold coupe.
        WinchM1Cmd.RunRequest := FALSE; WinchM1Cmd.ReqAscent := FALSE; WinchM1Cmd.ReqDescend := FALSE; WinchM1Cmd.StepTgt := 0;
        WinchM2Cmd.RunRequest := FALSE; WinchM2Cmd.ReqAscent := FALSE; WinchM2Cmd.ReqDescend := FALSE; WinchM2Cmd.StepTgt := 0;
        BucketCmd.ReqKoboldMeasureEnable := FALSE;

        TouchPositionM := M1_CablePosM;
        BottomTouched  := TRUE;   // variable d'info latchee (GEL AX8) - effacee a AX0 / AX_STAB / Reset
        IF LimitLegalDepthM < -0.01 THEN
            RaiseTargetM := MAX(TouchPositionM + RaiseOffBottomEff, LimitLegalDepthM + RaiseOffBottomEff);
        ELSE
            RaiseTargetM := TouchPositionM + RaiseOffBottomEff;
        END_IF;
        State := E_AutoCycleStep.AX9_RAISE_OFF_BOTTOM;

    E_AutoCycleStep.AX_DIVING_RETRY:
        CycleStep := E_AutoCycleStep.AX_DIVING_RETRY;
        CycleStateStr := 'AX_DIVING_RETRY - Reprise plongee : remonter au FDC haut';
        Lifecycle.Busy := TRUE;
        Lifecycle.Done := FALSE;
        ExpectedAxis := E_OperatorAxis.JOYSTICK_Y;
        ExpectedDirection := 1;
        WaitingForOperator := NOT JoystickDeflected;
        WaitingForProcess := JoystickDeflected;
        OperatorActionId := 16#0481;
        OperatorAction := 'AX_DIVING_RETRY - Reprise plongee : monter jusqu au FDC haut, puis relancer.';

        // Remontee assistee palier lent, Kobold coupe.
        WinchM1Cmd.RunRequest := CycleMotionPermit;
        WinchM1Cmd.ReqAscent := TRUE; WinchM1Cmd.ReqDescend := FALSE;
        WinchM1Cmd.StepTgt  := CST_StepSlow;
        WinchM2Cmd.RunRequest := CycleMotionPermit;
        WinchM2Cmd.ReqAscent := TRUE; WinchM2Cmd.ReqDescend := FALSE;
        WinchM2Cmd.StepTgt  := CST_StepSlow;
        BucketCmd.ReqKoboldMeasureEnable := FALSE;

        // AT-retry : treuils revenus au FDC haut -> nouvelle tentative de plongee.
        IF JoystickDeflected AND (WinchesAtTopWindow OR TopPositionSensor) THEN
            WinchM1Cmd.RunRequest := FALSE;
            WinchM2Cmd.RunRequest := FALSE;
            State := E_AutoCycleStep.AX4_DESCEND_DIVING;
        END_IF;

    (* ===================== EXTRACTION (AX9..AX12) ===================== *)

    E_AutoCycleStep.AX9_RAISE_OFF_BOTTOM:
        CycleStep := E_AutoCycleStep.AX9_RAISE_OFF_BOTTOM;
        CycleStateStr := 'AX9 - Retente les cables (palier 1), decollement du fond';
        Lifecycle.Busy := TRUE;
        Lifecycle.Done := FALSE;
        ExpectedAxis := E_OperatorAxis.JOYSTICK_Y;
        ExpectedDirection := 1;
        WaitingForOperator := NOT JoystickDeflected;
        WaitingForProcess := JoystickDeflected;
        OperatorActionId := 16#0409;
        OperatorAction := 'AX9 - Maintenir la montee palier 1 : retente des cables, decollement du fond.';

        // Palier 1 (doux). Selecteur couplage BOTH/M1/M2 = garde cote PRG_04 (GEL Q15),
        // le sequenceur commande toujours les deux treuils symetriquement.
        WinchM1Cmd.RunRequest := CycleMotionPermit;
        WinchM1Cmd.ReqAscent := TRUE; WinchM1Cmd.ReqDescend := FALSE;
        WinchM1Cmd.StepTgt := CST_StepSlow;
        WinchM2Cmd.RunRequest := CycleMotionPermit;
        WinchM2Cmd.ReqAscent := TRUE; WinchM2Cmd.ReqDescend := FALSE;
        WinchM2Cmd.StepTgt := CST_StepSlow;

        IF JoystickDeflected AND (M1_CablePosM >= RaiseTargetM) AND (M2_CablePosM >= RaiseTargetM) THEN
            WinchM1Cmd.RunRequest := FALSE;
            WinchM2Cmd.RunRequest := FALSE;
            State := E_AutoCycleStep.AX10_CLOSE_BUCKET;
        END_IF;

    E_AutoCycleStep.AX10_CLOSE_BUCKET:
        CycleStep := E_AutoCycleStep.AX10_CLOSE_BUCKET;
        CycleStateStr := 'AX10 - Fermeture benne (tolerance a peu pres ferme)';
        Lifecycle.Busy := TRUE;
        Lifecycle.Done := FALSE;
        ExpectedAxis := E_OperatorAxis.JOYSTICK_Y;
        ExpectedDirection := 1;
        WaitingForOperator := NOT JoystickDeflected;
        WaitingForProcess := JoystickDeflected;
        OperatorActionId := 16#040A;
        OperatorAction := 'AX10 - Maintenir la commande : fermeture de la benne.';

        // Etape benne seule : les DEUX treuils explicitement neutralises.
        WinchM1Cmd.RunRequest := FALSE; WinchM1Cmd.ReqAscent := FALSE; WinchM1Cmd.ReqDescend := FALSE; WinchM1Cmd.StepTgt := 0;
        WinchM2Cmd.RunRequest := FALSE; WinchM2Cmd.ReqAscent := FALSE; WinchM2Cmd.ReqDescend := FALSE; WinchM2Cmd.StepTgt := 0;
        BucketCmd.ReqClose := CycleMotionPermit;

        IF JoystickDeflected AND (Benne_Done AND (Benne_IsClosed OR Benne_IsRoughlyClosed)) THEN
            BucketCmd.ReqClose := FALSE;
            // C1e (GEL principe 4) : AX10 -> AX11 sans temps mort. M1+M2 lances le MEME
            // scan que la sortie AX10_CLOSE_BUCKET (pas de creux RunRequest a la frontiere).
            WinchM1Cmd.RunRequest := CycleMotionPermit;
            WinchM1Cmd.ReqAscent := TRUE; WinchM1Cmd.ReqDescend := FALSE;
            WinchM1Cmd.StepTgt  := CtrlAscentMaxStepEff;
            WinchM2Cmd.RunRequest := CycleMotionPermit;
            WinchM2Cmd.ReqAscent := TRUE; WinchM2Cmd.ReqDescend := FALSE;
            WinchM2Cmd.StepTgt  := CtrlAscentMaxStepEff;
            State := E_AutoCycleStep.AX11_CTRL_ASCENT;
        END_IF;

    E_AutoCycleStep.AX11_CTRL_ASCENT:
        CycleStep := E_AutoCycleStep.AX11_CTRL_ASCENT;
        CycleStateStr := 'AX11 - Remontee lente de controle';
        Lifecycle.Busy := TRUE;
        Lifecycle.Done := FALSE;
        ExpectedAxis := E_OperatorAxis.JOYSTICK_Y;
        ExpectedDirection := 1;
        WaitingForOperator := NOT JoystickDeflected;
        WaitingForProcess := JoystickDeflected;
        OperatorActionId := 16#040B;
        OperatorAction := 'AX11 - Maintenir la montee de controle : palier et synchronisme.';

        // Palier max reglable IHM, borne [1..2] (defaut 1 / P1 ; P2 possible au besoin).
        WinchM1Cmd.RunRequest := CycleMotionPermit;
        WinchM1Cmd.ReqAscent := TRUE; WinchM1Cmd.ReqDescend := FALSE;
        WinchM1Cmd.StepTgt  := CtrlAscentMaxStepEff;
        WinchM2Cmd.RunRequest := CycleMotionPermit;
        WinchM2Cmd.ReqAscent := TRUE; WinchM2Cmd.ReqDescend := FALSE;
        WinchM2Cmd.StepTgt  := CtrlAscentMaxStepEff;

        IF JoystickDeflected
           AND (M1_CablePosM >= (TouchPositionM + CtrlAscentDistM))
           AND (M2_CablePosM >= (TouchPositionM + CtrlAscentDistM))
           AND (ABS(M1_CablePosM - M2_CablePosM) <= CtrlAscentToleranceM) THEN
            State := E_AutoCycleStep.AX12_LOADED_ASCENT;
        END_IF;

    E_AutoCycleStep.AX12_LOADED_ASCENT:
        CycleStep := E_AutoCycleStep.AX12_LOADED_ASCENT;
        CycleStateStr := 'AX12 - Remontee en charge';
        Lifecycle.Busy := TRUE;
        Lifecycle.Done := FALSE;
        ExpectedAxis := E_OperatorAxis.JOYSTICK_Y;
        ExpectedDirection := 1;
        WaitingForOperator := NOT JoystickDeflected;
        WaitingForProcess := JoystickDeflected;
        OperatorActionId := 16#040C;
        OperatorAction := 'AX12 - Maintenir la montee en charge jusqu a la limite haute.';

        // Benne bien fermee -> palier 4 ; benne mal fermee (a peu pres) -> palier 1.
        // Pas de ralentissement 1 m avant la position top (montee franche).
        WinchM1Cmd.RunRequest := CycleMotionPermit;
        WinchM1Cmd.ReqAscent := TRUE; WinchM1Cmd.ReqDescend := FALSE;
        WinchM1Cmd.StepTgt  := SEL(Benne_IsClosed, CST_StepSlow, CST_StepLoaded);
        WinchM2Cmd.RunRequest := CycleMotionPermit;
        WinchM2Cmd.ReqAscent := TRUE; WinchM2Cmd.ReqDescend := FALSE;
        WinchM2Cmd.StepTgt  := SEL(Benne_IsClosed, CST_StepSlow, CST_StepLoaded);

        IF JoystickDeflected AND M1_CablePosM >= CableLimitM1AscentM THEN
            WinchM1Cmd.RunRequest := FALSE;
            WinchM2Cmd.RunRequest := FALSE;
            State := E_AutoCycleStep.AX13_DRAIN_PAUSE;
        END_IF;

    (* ===================== DECHARGE (AX13..AX18) ===================== *)

    E_AutoCycleStep.AX13_DRAIN_PAUSE:
        CycleStep := E_AutoCycleStep.AX13_DRAIN_PAUSE;
        CycleStateStr := 'AX13 - Egouttage du godet en cours';
        Lifecycle.Busy := TRUE;
        Lifecycle.Done := FALSE;
        ExpectedAxis := E_OperatorAxis.NONE;
        ExpectedDirection := 0;
        WaitingForOperator := FALSE;
        WaitingForProcess := TRUE;
        OperatorActionId := 16#0409;
        OperatorAction := 'AX13 - Egouttage : attendre la tempo ou appuyer sur "passer egouttage".';
        WinchM1Cmd.RunRequest := FALSE;
        WinchM2Cmd.RunRequest := FALSE;

        // Tempo d'egouttage armee/remise a zero en §1 (gate sur State = AX13, PT = DrainTimeEff).
        // Duree reglable IHM (CfgDrainTime) + bypass immediat (SkipDrainEdge).
        IF JoystickDeflected AND (DrainingTimer.Q OR SkipDrainEdge.Q) THEN
            State := E_AutoCycleStep.AX14_TRANSLATE_DUMP;
        END_IF;

    E_AutoCycleStep.AX14_TRANSLATE_DUMP:
        CycleStep := E_AutoCycleStep.AX14_TRANSLATE_DUMP;
        CycleStateStr := 'AX14 - Deplacement vers tremie (grille/crible libres)';
        Lifecycle.Busy := TRUE;
        Lifecycle.Done := FALSE;
        ExpectedAxis := E_OperatorAxis.JOYSTICK_X;
        ExpectedDirection := -1;
        WaitingForOperator := NOT JoystickDeflected;
        WaitingForProcess := JoystickDeflected;
        OperatorActionId := 16#040A;
        OperatorAction := 'AX14 - Maintenir la translation vers la tremie de dechargement.';

        TranslationCmd.PositionTgt := 1; // Trémie
        TranslationCmd.ReqStart := CycleMotionPermit;

        IF JoystickDeflected AND Translation_At_Tremie THEN
            TranslationCmd.ReqStart := FALSE;
            State := E_AutoCycleStep.AX15A_DUMP_ARRIVE;
        END_IF;

    E_AutoCycleStep.AX15A_DUMP_ARRIVE:
        CycleStep := E_AutoCycleStep.AX15A_DUMP_ARRIVE;
        CycleStateStr := 'AX15a - Arrivee tremie : treuils arretes, attente ouverture';
        Lifecycle.Busy := TRUE;
        Lifecycle.Done := FALSE;
        ExpectedAxis := E_OperatorAxis.JOYSTICK_Y;
        ExpectedDirection := -1;
        WaitingForOperator := NOT JoystickDeflected;
        WaitingForProcess := JoystickDeflected;
        OperatorActionId := 16#040B;
        OperatorAction := 'AX15a - A la tremie : deflechir vers le bas pour ouvrir la benne et vider.';

        // Config treuil UNIQUE : arret des deux treuils (aucune descente couplee ici).
        WinchM1Cmd.RunRequest := FALSE; WinchM1Cmd.ReqAscent := FALSE; WinchM1Cmd.ReqDescend := FALSE; WinchM1Cmd.StepTgt := 0;
        WinchM2Cmd.RunRequest := FALSE; WinchM2Cmd.ReqAscent := FALSE; WinchM2Cmd.ReqDescend := FALSE; WinchM2Cmd.StepTgt := 0;

        // Geste operateur (manche defleci) -> phase d'ouverture benne.
        IF JoystickDeflected THEN
            State := E_AutoCycleStep.AX15B_DUMP_OPEN;
        END_IF;

    E_AutoCycleStep.AX15B_DUMP_OPEN:
        CycleStep := E_AutoCycleStep.AX15B_DUMP_OPEN;
        CycleStateStr := 'AX15b - Vidage : ouverture benne pour vider le contenu, treuils arretes';
        Lifecycle.Busy := TRUE;
        Lifecycle.Done := FALSE;
        ExpectedAxis := E_OperatorAxis.JOYSTICK_Y;
        ExpectedDirection := -1;
        WaitingForOperator := NOT JoystickDeflected;
        WaitingForProcess := JoystickDeflected;
        OperatorActionId := 16#040B;
        OperatorAction := 'AX15b - Maintenir : ouverture complete de la benne, vidage a la tremie.';

        // Config treuil UNIQUE : etape benne seule, les deux treuils neutralises
        // (plus de descente couplee M1+M2 simultanee a l'ouverture benne -> plus
        // d'ecart M1/M2 volontaire ni de faux SafeStop concordance contacteurs).
        WinchM1Cmd.RunRequest := FALSE; WinchM1Cmd.ReqAscent := FALSE; WinchM1Cmd.ReqDescend := FALSE; WinchM1Cmd.StepTgt := 0;
        WinchM2Cmd.RunRequest := FALSE; WinchM2Cmd.ReqAscent := FALSE; WinchM2Cmd.ReqDescend := FALSE; WinchM2Cmd.StepTgt := 0;

        BucketCmd.ReqOpen := CycleMotionPermit;

        // Option operateur (bit IHM) : descendre la benne dans la gueule de tremie
        // pour aider la vidange -> repositionnement couple M1+M2 (AX15C). Prioritaire
        // sur la fin de vidage.
        IF RepositionRequest THEN
            State := E_AutoCycleStep.AX15C_DUMP_REPOSITION;
        ELSIF JoystickDeflected AND Benne_Done AND Benne_IsOpen THEN
            BucketCmd.ReqOpen := FALSE;
            State := E_AutoCycleStep.AX18_DONE_SYNC;
        END_IF;

    E_AutoCycleStep.AX15C_DUMP_REPOSITION:
        CycleStep := E_AutoCycleStep.AX15C_DUMP_REPOSITION;
        CycleStateStr := 'AX15c - Repositionnement couple M1+M2 (aide vidange tremie)';
        Lifecycle.Busy := TRUE;
        Lifecycle.Done := FALSE;
        ExpectedAxis := E_OperatorAxis.JOYSTICK_Y;
        ExpectedDirection := -1;
        WaitingForOperator := NOT JoystickDeflected;
        WaitingForProcess := JoystickDeflected;
        OperatorActionId := 16#040C;
        OperatorAction := 'AX15c - Descente couplee M1+M2 ; relacher l option pour reprendre le vidage.';

        // Descente couplee M1+M2, palier lent, sous homme-mort. Commandes SYMETRIQUES
        // (meme sens, meme palier) -> FB_SyncDeviation actif, pas d'ecart volontaire.
        WinchM1Cmd.ReqAscent := FALSE; WinchM1Cmd.ReqDescend := TRUE;
        WinchM1Cmd.RunRequest := CycleMotionPermit;
        WinchM1Cmd.StepTgt := CST_StepSlow;
        WinchM2Cmd.ReqAscent := FALSE; WinchM2Cmd.ReqDescend := TRUE;
        WinchM2Cmd.RunRequest := CycleMotionPermit;
        WinchM2Cmd.StepTgt := CST_StepSlow;

        // La benne reste ouverte pendant le repositionnement (on finit l'ouverture si besoin).
        BucketCmd.ReqOpen := CycleMotionPermit AND NOT Benne_IsOpen;

        // Retour a AX15B des que l'operateur relache l'option de repositionnement.
        IF NOT RepositionRequest THEN
            WinchM1Cmd.RunRequest := FALSE;
            WinchM2Cmd.RunRequest := FALSE;
            State := E_AutoCycleStep.AX15B_DUMP_OPEN;
        END_IF;

    E_AutoCycleStep.AX18_DONE_SYNC:
        CycleStep := E_AutoCycleStep.AX18_DONE_SYNC;
        CycleStateStr := 'AX18 - Passe terminee : aller en P1 pour recommencer';
        WinchM1Cmd.RunRequest := FALSE;
        WinchM2Cmd.RunRequest := FALSE;
        TranslationCmd.ReqStart := FALSE;
        Lifecycle.Done := TRUE;
        Lifecycle.Busy := FALSE;
        ExpectedAxis := E_OperatorAxis.JOYSTICK_X;
        ExpectedDirection := 1;
        WaitingForOperator := TRUE;
        WaitingForProcess := FALSE;
        OperatorActionId := 16#040D;
        OperatorAction := 'AX18 - Cycle termine. Aller en P1 (joystick vers la droite) pour recommencer.';

        // Compteur de prélèvements (RETAIN) + durée du cycle — F2: cadré par front (1 seul par cycle)
        IF NOT SampleCountDone THEN
            SampleCount := SampleCount + 1;
            LastCycleDuration := CurrentCycleElapsed;   // fige la durée du cycle qui vient de s'achever
            SampleCountDone := TRUE;
        END_IF;

        // Rebouclage DIRECT sur AX2_TRANSLATE_P1 (GEL Q14) : la machine est deja
        // referencee, la passe suivante enchaine sur la translation P1 (pas de retour AX0).
        // Relance sur StartCycle OU FRONT joystick (geste franc) - pas sur simple maintien,
        // pour que AX18 (Lifecycle.Done + msg) soit reellement observable / tracable.
        IF StartEdge.Q OR JoyDeflectedEdge.Q THEN
            SampleCountDone := FALSE;
            Lifecycle.Done := FALSE;
            State := E_AutoCycleStep.AX2_TRANSLATE_P1;
        END_IF;

    E_AutoCycleStep.AX_STAB:
        CycleStep := E_AutoCycleStep.AX_STAB;
        CycleStateStr := 'AX_STAB - Cycle en attente / stabilisation sur anomalie';
        WinchM1Cmd.RunRequest := FALSE; WinchM1Cmd.ReqAscent := FALSE; WinchM1Cmd.ReqDescend := FALSE;
        WinchM2Cmd.RunRequest := FALSE; WinchM2Cmd.ReqAscent := FALSE; WinchM2Cmd.ReqDescend := FALSE;
        TranslationCmd.ReqStart := FALSE;
        BucketCmd.ReqOpen := FALSE;
        BucketCmd.ReqClose := FALSE;
        BucketCmd.ReqKoboldMeasureEnable := FALSE;   // Coupure contacteur Kobold au repli defaut (0 ordre residuel)
        Lifecycle.Busy := FALSE;
        Lifecycle.Done := FALSE;
        ExpectedAxis := E_OperatorAxis.BUTTON;
        ExpectedDirection := 0;
        WaitingForOperator := TRUE;
        WaitingForProcess := FALSE;
        OperatorActionId := 16#0480;
        OperatorAction := 'AX_STAB - Cycle stabilise sur anomalie : acquitter le defaut pour reinitialiser.';

END_CASE;
END_IF;
{endregion}

{region "§4 Repli homme mort & Syntheses"}
// 🛑 Relâchement du manche (retour au centre) OU de l'homme-mort : neutralisation
// des demandes actives. Gate continu : aucune commande d'actionneur ne survit à la
// perte du permis opérateur (manche défléchi ET homme-mort armé).
IF Lifecycle.Busy AND NOT CycleMotionPermit THEN
    WinchM1Cmd.RunRequest := FALSE;
    WinchM2Cmd.RunRequest := FALSE;
    TranslationCmd.ReqStart := FALSE;
    BucketCmd.ReqOpen := FALSE;
    BucketCmd.ReqClose := FALSE;
    BucketCmd.ReqKoboldMeasureEnable := FALSE;
END_IF;

RequestActive := WinchM1Cmd.RunRequest OR WinchM2Cmd.RunRequest OR TranslationCmd.ReqStart OR BucketCmd.ReqOpen OR BucketCmd.ReqClose OR BucketCmd.ReqKoboldMeasureEnable; // Somme logique complete des demandes (contacteur Kobold inclus)
{endregion}

END_FUNCTION_BLOCK

(* ---- FB_DiveSearch.st ---- *)
(* =======================================================================
   FB_DiveSearch - Assistance plongee et recherche du fond Kobold
   Role : qualifier l'immersion et autoriser la descente assistee.
   Interface : contrat standard + bus Inputs/Outputs.
   Documentation : DOC/AF/AF_Partie-04_Mode_SemiAuto_Sequenceur_v2.3.md
   ======================================================================= *)
FUNCTION_BLOCK FB_DiveSearch
VAR_INPUT
    // === CONTRAT STANDARD ===
    Enable                  : BOOL;                   // --> [CMD] Autorisation generale du FB
    Reset                   : BOOL;                   // --> [CMD] Acquittement defaut sur front

    // === BUS FONCTIONNEL ===
    Inputs                  : ST_fbDiveSearch_Inputs; // --> [BUS] Commande, capteurs et reglages
END_VAR
VAR_OUTPUT
    // === STATUT IEC ===
    Ready                   : BOOL;                   // <-- [STAT] FB pret a fonctionner
    Fault                   : ST_Fault;               // <-- [DIAG] Defaut live et latche
    Lifecycle               : ST_Lifecycle;           // <-- [STAT] Cycle en cours / termine

    // === BUS FONCTIONNEL ===
    Outputs                 : ST_fbDiveSearch_Outputs;// <-- [BUS] Etat, permis et diagnostic
END_VAR
VAR
    // === SOUS-INSTANCES & FRONTS ===
    ResetEdge               : R_TRIG;                 // . [LOC] Front Reset
    ErrorEdge               : R_TRIG;                 // . [LOC] Apparition d'un defaut
    KoboldRiseEdge          : R_TRIG;                 // . [LOC] Entree dans l'eau
    KoboldFallEdge          : F_TRIG;                 // . [LOC] Sortie de l'eau / fond
    instFault               : FB_FaultCore;           // * [INST] Socle defaut transverse
    instCauses              : ARRAY[0..15] OF ST_FaultCause; // . [LOC] Causes nommees

    // === CALCULS DE GARDE ===
    ImmersionCourse_M          : REAL;                // . [LOC] Course maximale vers immersion (m)
    BottomCourse_M             : REAL;                // . [LOC] Course maximale vers fond (m)
    CalculatedImmersionTimeout : TIME;                // . [LOC] Timeout immersion calcule
    CalculatedBottomTimeout    : TIME;                // . [LOC] Timeout fond calcule
    EffectiveDiveSpeedMin_Mps  : REAL;                // . [LOC] Vitesse minimale appliquee (m/s)
    EffectiveTimeoutMargin     : REAL;                // . [LOC] Marge appliquee au calcul
    EffectiveTimeoutMinCourse_M: REAL;                // . [LOC] Plancher de course applique (m)
    EffectiveTimeoutMaxCourse_M: REAL;                // . [LOC] Plafond de course applique (m)
    EffectiveSecToMs            : REAL;               // . [LOC] Conversion secondes/millisecondes

    // === MEMORISATIONS & TEMPORISATIONS ===
    ImmersionTimerAcc       : TIME := T#0ms;          // . [LOC] Temps effectif de recherche immersion
    BottomTimerAcc          : TIME := T#0ms;          // . [LOC] Temps effectif de recherche fond
    PrevState               : E_DiveSearchState;      // . [LOC] Etat du scan precedent
    ImmersionConfirmed      : BOOL;                   // . [LOC] Immersion validee
    StepAtFaultCaptured     : BOOL;                   // . [LOC] Etape de defaut deja figee

    // === CAUSES INTERNES ===
    ErrorCausePresent       : BOOL;                   // . [LOC] Parametrage invalide
    SeqErrorFault           : BOOL;                   // . [LOC] Incoherence de sequence
    Palier5ForbiddenFault   : BOOL;                   // . [LOC] Palier 5 interdit sous Kobold
    TimeoutImmersionFault   : BOOL;                   // . [LOC] Timeout recherche immersion
    TimeoutBottomFault      : BOOL;                   // . [LOC] Timeout recherche fond
    DescentActive           : BOOL;                   // . [LOC] Descending demandee et autorisee
END_VAR

{region "§1 Fronts, calculs et causes"}
ResetEdge(CLK := Reset);
KoboldRiseEdge(CLK := Inputs.KoboldImmersed);
KoboldFallEdge(CLK := Inputs.KoboldImmersed);

// Les valeurs par defaut du DUT couvrent l'appel sans configuration explicite.
// Le repli runtime protege aussi un appel avec une structure entierement nulle.
EffectiveDiveSpeedMin_Mps := Inputs.Config.DiveSpeedMin_Mps;
IF EffectiveDiveSpeedMin_Mps <= 0.0 THEN EffectiveDiveSpeedMin_Mps := 0.15; END_IF;
EffectiveTimeoutMargin := Inputs.Config.TimeoutMarginFactor;
IF EffectiveTimeoutMargin <= 0.0 THEN EffectiveTimeoutMargin := 1.5; END_IF;
EffectiveTimeoutMinCourse_M := Inputs.Config.TimeoutMinCourse_M;
IF EffectiveTimeoutMinCourse_M <= 0.0 THEN EffectiveTimeoutMinCourse_M := 1.0; END_IF;
EffectiveTimeoutMaxCourse_M := Inputs.Config.TimeoutMaxCourse_M;
IF EffectiveTimeoutMaxCourse_M < EffectiveTimeoutMinCourse_M THEN EffectiveTimeoutMaxCourse_M := 200.0; END_IF;
EffectiveSecToMs := Inputs.Config.SecToMs;
IF EffectiveSecToMs <= 0.0 THEN EffectiveSecToMs := 1000.0; END_IF;

ErrorCausePresent := (Inputs.CycleTime <= T#0ms)
                 OR (NOT Inputs.BypassPreconditions AND (
                       (Inputs.DiveStartMin_M < Inputs.ImmersionUpper_M)
                    OR (Inputs.ImmersionUpper_M <= Inputs.ImmersionLower_M)
                    OR (Inputs.ImmersionLower_M <= Inputs.LimitLegalDepthMin_M)
                    OR (Inputs.CableLimitAscent_M <= Inputs.ImmersionLower_M)));

ImmersionCourse_M := LIMIT(EffectiveTimeoutMinCourse_M,
                           Inputs.CableLimitAscent_M - Inputs.ImmersionLower_M,
                           EffectiveTimeoutMaxCourse_M);
BottomCourse_M := LIMIT(EffectiveTimeoutMinCourse_M,
                        Inputs.ImmersionLower_M - Inputs.LimitLegalDepthMin_M,
                        EffectiveTimeoutMaxCourse_M);
CalculatedImmersionTimeout := UDINT_TO_TIME(REAL_TO_UDINT(
    ImmersionCourse_M / EffectiveDiveSpeedMin_Mps * EffectiveTimeoutMargin * EffectiveSecToMs));
CalculatedBottomTimeout := UDINT_TO_TIME(REAL_TO_UDINT(
    BottomCourse_M / EffectiveDiveSpeedMin_Mps * EffectiveTimeoutMargin * EffectiveSecToMs));

IF (Outputs.StepState = E_DiveSearchState.SEARCHING_IMMERSION)
   AND Inputs.MotionRequestActive AND (Inputs.MotionDirection = -1) THEN
    ImmersionTimerAcc := ImmersionTimerAcc + Inputs.CycleTime;
    IF ImmersionTimerAcc >= CalculatedImmersionTimeout THEN TimeoutImmersionFault := TRUE; END_IF;
END_IF;

IF (Outputs.StepState = E_DiveSearchState.SEARCHING_BOTTOM)
   AND Inputs.MotionRequestActive AND (Inputs.MotionDirection = -1) THEN
    BottomTimerAcc := BottomTimerAcc + Inputs.CycleTime;
    IF BottomTimerAcc >= CalculatedBottomTimeout THEN TimeoutBottomFault := TRUE; END_IF;
END_IF;

IF ResetEdge.Q AND NOT ErrorCausePresent AND NOT Inputs.KoboldImmersed
   AND NOT Inputs.MotionRequestActive AND NOT (Inputs.CurrentSpeedStep > 4) THEN
    SeqErrorFault := FALSE;
    Palier5ForbiddenFault := FALSE;
    TimeoutImmersionFault := FALSE;
    TimeoutBottomFault := FALSE;
    ImmersionTimerAcc := T#0ms;
    BottomTimerAcc := T#0ms;
    ImmersionConfirmed := FALSE;
    Outputs.BottomTouchConfirmed := FALSE;
    Outputs.StepAtFault := E_DiveSearchState.WAIT_PRECONDITIONS;
    StepAtFaultCaptured := FALSE;
    Outputs.StepState := E_DiveSearchState.WAIT_PRECONDITIONS;
END_IF;

instCauses[0].Active := SeqErrorFault;
instCauses[0].Latching := TRUE;
instCauses[0].Texte := 'Incoherence sequence immersion Kobold';
instCauses[1].Active := ErrorCausePresent;
instCauses[1].Latching := TRUE;
instCauses[1].Texte := 'Parametrage invalide des seuils de plongee';
instCauses[2].Active := Palier5ForbiddenFault;
instCauses[2].Latching := TRUE;
instCauses[2].Texte := 'Palier 5 interdit pendant la mesure Kobold';
instCauses[3].Active := TimeoutImmersionFault;
instCauses[3].Latching := TRUE;
instCauses[3].Texte := 'Timeout recherche immersion Kobold';
instCauses[4].Active := TimeoutBottomFault;
instCauses[4].Latching := TRUE;
instCauses[4].Texte := 'Timeout recherche fond Kobold';

instFault(Enable := Enable, Reset := Reset, Causes := instCauses);
Fault := instFault.Fault;

ErrorEdge(CLK := Fault.Error);
IF ErrorEdge.Q AND NOT StepAtFaultCaptured THEN
    Outputs.StepAtFault := PrevState;
    StepAtFaultCaptured := TRUE;
ELSIF ResetEdge.Q AND NOT ErrorCausePresent AND NOT Inputs.KoboldImmersed
      AND NOT Inputs.MotionRequestActive AND NOT (Inputs.CurrentSpeedStep > 4) THEN
    Outputs.StepAtFault := E_DiveSearchState.WAIT_PRECONDITIONS;
END_IF;
{endregion}

{region "§2 Neutralisation et machine d'etat"}
IF NOT Enable OR NOT Inputs.PowerContactorEngaged THEN
    Ready := FALSE;
    Lifecycle.Busy := FALSE;
    Lifecycle.Done := FALSE;
    Outputs.DescendPermit := FALSE;
    Outputs.KoboldContactorCmd := FALSE;
    Outputs.BottomTouchConfirmed := FALSE;
    Outputs.StepState := E_DiveSearchState.WAIT_PRECONDITIONS;
    Outputs.OperatorActionId := 0;
    Outputs.OperatorAction := '';
    ImmersionConfirmed := FALSE;
    ImmersionTimerAcc := T#0ms;
    BottomTimerAcc := T#0ms;
    Outputs.MinStepDown := 0;
    PrevState := E_DiveSearchState.WAIT_PRECONDITIONS;
    RETURN;
END_IF;

Ready := Enable AND NOT Fault.Latched;
Outputs.DescendPermit := FALSE;
Outputs.KoboldContactorCmd := FALSE;
Lifecycle.Busy := FALSE;
Lifecycle.Done := FALSE;
Outputs.OperatorActionId := 0;
Outputs.OperatorAction := '';

DescentActive := Inputs.MotionRequestActive AND (Inputs.MotionDirection = -1)
              AND ((Inputs.Mode = E_Mode.MAINT_N1) OR (Inputs.Mode = E_Mode.MAINT_N2))
              AND NOT (Inputs.CurrentSpeedStep > 4)
              AND NOT SeqErrorFault;

IF Fault.Error OR Fault.Latched THEN
    Outputs.StepState := E_DiveSearchState.ERROR_HOLD;
    Outputs.KoboldContactorCmd := FALSE;
    Outputs.OperatorActionId := 16#0180;
    Outputs.OperatorAction := 'Verifier les conditions puis rearmer avant une nouvelle plongee.';
ELSE
    CASE Outputs.StepState OF
        E_DiveSearchState.WAIT_PRECONDITIONS:
            IF NOT Inputs.BypassPreconditions
               AND (NOT Inputs.BucketIsOpen OR NOT Inputs.PositionsValid OR Inputs.KoboldImmersed
                    OR (Inputs.M1Position_M < Inputs.DiveStartMin_M)
                    OR (Inputs.M2Position_M < Inputs.DiveStartMin_M)) THEN
                Outputs.OperatorActionId := 16#0100;
                Outputs.OperatorAction := 'Verifier benne ouverte, positions et Kobold au repos.';
            ELSE
                Outputs.StepState := E_DiveSearchState.READY_TO_DESCEND;
            END_IF;

        E_DiveSearchState.READY_TO_DESCEND:
            Ready := TRUE;
            Outputs.OperatorActionId := 16#0101;
            Outputs.OperatorAction := 'Demander une descente pour rechercher le fond.';
            IF Inputs.MotionRequestActive AND (Inputs.MotionDirection = -1) THEN
                ImmersionTimerAcc := T#0ms;
                Outputs.StepState := E_DiveSearchState.SEARCHING_IMMERSION;
            END_IF;

        E_DiveSearchState.SEARCHING_IMMERSION:
            Lifecycle.Busy := TRUE;
            Outputs.DescendPermit := DescentActive;
            Outputs.KoboldContactorCmd := DescentActive;
            Outputs.OperatorActionId := 16#0102;
            Outputs.OperatorAction := 'Maintenir la descente : recherche immersion Kobold.';
            IF Inputs.CurrentSpeedStep > 4 THEN
                IF NOT StepAtFaultCaptured THEN
                    Outputs.StepAtFault := Outputs.StepState;
                    StepAtFaultCaptured := TRUE;
                END_IF;
                Palier5ForbiddenFault := TRUE;
            END_IF;
            IF KoboldRiseEdge.Q THEN
                IF (Inputs.M1Position_M <= Inputs.ImmersionUpper_M)
                   AND (Inputs.M1Position_M >= Inputs.ImmersionLower_M)
                   AND (Inputs.M2Position_M <= Inputs.ImmersionUpper_M)
                   AND (Inputs.M2Position_M >= Inputs.ImmersionLower_M) THEN
                    ImmersionConfirmed := TRUE;
                    BottomTimerAcc := T#0ms;
                    Outputs.StepState := E_DiveSearchState.SEARCHING_BOTTOM;
                ELSE
                    IF NOT StepAtFaultCaptured THEN
                        Outputs.StepAtFault := Outputs.StepState;
                        StepAtFaultCaptured := TRUE;
                    END_IF;
                    SeqErrorFault := TRUE;
                END_IF;
            ELSIF (Inputs.M1Position_M < Inputs.ImmersionLower_M)
               OR (Inputs.M2Position_M < Inputs.ImmersionLower_M) THEN
                IF NOT StepAtFaultCaptured THEN
                    Outputs.StepAtFault := Outputs.StepState;
                    StepAtFaultCaptured := TRUE;
                END_IF;
                SeqErrorFault := TRUE;
            END_IF;

        E_DiveSearchState.SEARCHING_BOTTOM:
            Lifecycle.Busy := TRUE;
            Outputs.DescendPermit := DescentActive;
            Outputs.KoboldContactorCmd := DescentActive;
            Outputs.OperatorActionId := 16#0103;
            Outputs.OperatorAction := 'Maintenir la descente : immersion validee, recherche du fond.';
            IF Inputs.CurrentSpeedStep > 4 THEN
                IF NOT StepAtFaultCaptured THEN
                    Outputs.StepAtFault := Outputs.StepState;
                    StepAtFaultCaptured := TRUE;
                END_IF;
                Palier5ForbiddenFault := TRUE;
            END_IF;
            IF KoboldFallEdge.Q AND ImmersionConfirmed THEN
                Outputs.BottomTouchConfirmed := TRUE;
                ImmersionConfirmed := FALSE;
                Outputs.KoboldContactorCmd := FALSE;
                Outputs.StepState := E_DiveSearchState.BOTTOM_CONFIRMED;
            END_IF;

        E_DiveSearchState.BOTTOM_CONFIRMED:
            Lifecycle.Done := TRUE;
            Outputs.KoboldContactorCmd := FALSE;
            Outputs.OperatorActionId := 16#0104;
            Outputs.OperatorAction := 'Fond detecte : demander la fermeture ou extraction.';

        E_DiveSearchState.ERROR_HOLD:
            Outputs.KoboldContactorCmd := FALSE;
    END_CASE;
END_IF;

IF DescentActive AND ((Outputs.StepState = E_DiveSearchState.SEARCHING_IMMERSION)
                   OR (Outputs.StepState = E_DiveSearchState.SEARCHING_BOTTOM)) THEN
    Outputs.MinStepDown := LIMIT(0, Inputs.CfgDiveFloorStep, 5);
ELSE
    Outputs.MinStepDown := 0;
END_IF;

PrevState := Outputs.StepState;
{endregion}

END_FUNCTION_BLOCK

(* ---- FB_ExtractionAssist.st ---- *)
(* =======================================================================
   ⚙️ FB_ExtractionAssist — Fermeture benne et remontée assistée
   ───────────────────────────────────────────────────────────────
   🎯 Rôle : Séquence d'extraction (fermeture benne, remontée de contrôle, remontée nominale)
   🛡️ Sécurité : Aucune remontée assistée sans fond confirmé, contrôle palier 1
   📄 Doc métier : DOC/AF/AF_Partie-04_Mode_SemiAuto_Sequenceur_v2.3.md
   ======================================================================= *)
FUNCTION_BLOCK FB_ExtractionAssist
VAR_INPUT
    // === COMMANDES & AUTORISATIONS ===
    Enable                      : BOOL;     // --> [CMD] Activation generale du FB (TRUE=Autorise)
    Reset                       : BOOL;     // --> [CMD] Acquittement defaut (front)
    PowerContactorEngaged       : BOOL;     // --> [SAFE] Chaine de securite OK
    Mode                        : E_Mode;   // --> [CMD] Mode de fonctionnement arbitre
    MotionRequestActive         : BOOL;     // --> [CMD] Intention de mouvement active
    MotionDirection             : INT;      // --> [CMD] Sens de mouvement (+1 = montee)
    BottomPositionConfirmed     : BOOL;     // --> [SAFE] Attestation fond confirme (Kobold ou op)

    // === CAPTEURS & ETATS MATERIELS ===
    BucketIsClosed              : BOOL;     // --> [HW] Benne fermee confirmee
    BucketBusy                  : BOOL;     // --> [HW] Mouvement benne en cours
    BucketError                 : BOOL;     // --> [SAFE] Defaut sur sous-systeme benne
    WinchSyncError              : BOOL;     // --> [SAFE] Defaut de desynchronisme treuils M1/M2
    M1Position_M                : REAL;     // --> [HW] Position codeur treuil M1 (m)
    M2Position_M                : REAL;     // --> [HW] Position codeur treuil M2 (m)
    M1MeasuredSpeedValid        : BOOL;     // --> [HW] Validite mesure vitesse M1
    M2MeasuredSpeedValid        : BOOL;     // --> [HW] Validite mesure vitesse M2
    PositionsValid              : BOOL;     // --> [HW] Validite des mesures de position

    // === CONFIGURATION & REGLAGES ===
    ControlAscentDistance_M     : REAL;     // --> [CFG] Distance palier 1 de controle remontee (m)
    CfgBucketCloseTimeout       : TIME := T#75s;// --> [CFG] Backstop fermeture benne (doit rester > BucketMoveTimeout)
    BucketMoveTimeout           : TIME := T#60s;// --> [CFG] Reference watchdog mouvement FB_Bucket (verrouillage ordre backstop)
    CycleTime                   : TIME := T#10ms;// --> [CFG] Base de temps d'integration (periode MainTask)
END_VAR
VAR_OUTPUT
    // === ETATS IEC & DEFECTUOSITES ===
    Ready                       : BOOL;     // <-- [STAT] FB pret a fonctionner
    // 🧩 Statut transverse (forme cible ST_Fault + ST_Lifecycle)
    Fault                       : ST_Fault;
    Lifecycle                   : ST_Lifecycle;
    ExtractionState             : E_ExtractionAssistState; // <-- [STAT] Phase interne extraction
    StepAtFault                 : E_ExtractionAssistState; // <-- [DIAG] Phase active memorisee lors du defaut

    // === ORDRES & AUTORISATIONS ===
    BucketCloseRequest          : BOOL;     // <-- [ACT] Demande de fermeture benne
    AscentPermit                : BOOL;     // <-- [ACT] Autorisation de remontee assistee
    ExtractionControlActive     : BOOL;     // <-- [ACT] Plafond palier 1 pendant la montee controlee
    BottomConfirmationConsumed  : BOOL;     // <-- [STAT] Signal confirmation fond consomme

    // === DIAGNOSTIC IHM ===
    OperatorActionId            : WORD;     // <-- [DIAG] ID action operateur requise
    OperatorAction              : STRING(120); // <-- [DIAG] Message explicatif operateur
END_VAR
VAR
    // === DETECTEURS DE FRONTS ===
    ResetEdge                   : R_TRIG;   // . [LOC] Detecteur front montant Reset
    ErrorEdge                   : R_TRIG;   // . [LOC] Detecteur front montant apparition defaut

    // === MEMORISATIONS & POSITIONS INTERNES ===
    ControlStartM1Position_M    : REAL;     // . [LOC] Position M1 au debut du palier de controle (m)
    ControlStartM2Position_M    : REAL;     // . [LOC] Position M2 au debut du palier de controle (m)
    PrevState                   : E_ExtractionAssistState; // . [LOC] Phase au scan precedent (survit au gate)

    // === CALCUL DYNAMIQUE RUNTIME DU TIMEOUT DECOLLAGE ===
    CalculatedControlAscentTimeout : TIME;  // . [LOC] Plafond anti-blocage decollage calcule au runtime

    // === ACCUMULATEURS DE TEMPS ANTI-POMPAGE ===
    BucketCloseTimerAcc         : TIME := T#0ms;// . [LOC] Temps cumule fermeture benne sous montee demandee
    ControlAscentTimerAcc       : TIME := T#0ms;// . [LOC] Temps cumule decollage controle sous montee demandee

    // === VARIABLES LOCALES INTERNES ===
    ErrorCausePresent           : BOOL;     // . [LOC] Presence d'une cause de defaut parametrage
    BucketErrorFault            : BOOL;     // . [LOC] Latch erreur benne
    SyncOrSpeedErrorFault       : BOOL;     // . [LOC] Latch erreur synchro/vitesse
    TimeoutBucketCloseFault     : BOOL;     // . [LOC] Latch backstop fermeture benne
    TimeoutControlAscentFault   : BOOL;     // . [LOC] Latch timeout decollage controle
    StepAtFaultCaptured         : BOOL;     // . [LOC] StepAtFault deja fige pour l'episode de defaut courant
    AssistPermit                : BOOL;     // . [LOC] Ascending assistee reellement demandee (sens + mode)
    AscentControlSafe           : BOOL;     // . [LOC] Entrees [SAFE] saines pour le decollage controle
    AscentNominalSafe           : BOOL;     // . [LOC] Entrees [SAFE] saines pour la remontee nominale
    CausesPhysiquesEffacees     : BOOL;     // . [LOC] Toutes les entrees defaut treuil/benne revenues a l'etat sain

    // === SOCLE DEFAUT ===
    instFault                   : FB_FaultCore;                  // * [INST] Socle défaut transverse
    instCauses                  : ARRAY[0..15] OF ST_FaultCause; // . [LOC] Table des causes nommées
END_VAR
VAR CONSTANT
    // === CONSTANTES DERIVATION TIMEOUT ANTI-BLOCAGE ===
    CST_MinSpeed_Mps            : REAL := 0.15;   // Vitesse Palier 1 mini sous charge/mou (m/s)
    CST_ControlAscentMargin     : REAL := 2.0;    // Facteur de marge sur la course de decollage
    CST_TimeoutMinDistance_M    : REAL := 0.1;    // Plancher de distance pour le calcul (evite timeout degenere)
    CST_TimeoutMaxDistance_M    : REAL := 20.0;   // Plafond de distance : borne le calcul avant REAL_TO_UDINT (anti-overflow)
    CST_BackstopMax             : TIME := T#600s; // Plafond du backstop fermeture benne : au-dela, risque d'overflow de l'accumulateur
    CST_SecToMs                 : REAL := 1000.0; // Conversion secondes -> millisecondes
END_VAR

// === IMPLEMENTATION ===

{region "§1 Causes & Socle Défaut (évalué en continu)"}
// 🔑 1. FRONTS
ResetEdge(CLK := Reset);
// Parametrage invalide : distance nulle, backstop nul, base de temps nulle, ou backstop
// qui fauterait AVANT le watchdog benne (masquerait BucketError - ordre des watchdogs).
ErrorCausePresent := (ControlAscentDistance_M <= 0.0)
                  OR (CfgBucketCloseTimeout <= T#0ms)
                  OR (CycleTime <= T#0ms)
                  OR (CfgBucketCloseTimeout <= BucketMoveTimeout)
                  OR (CfgBucketCloseTimeout > CST_BackstopMax);  // borne haute : evite l'overflow de BucketCloseTimerAcc (F3)

// ⏱️ Plafond anti-blocage decollage calcule au runtime : course de controle bornee [plancher..plafond]
// avant conversion REAL->UDINT->TIME (anti-overflow sur valeur IHM aberrante, CQS §6).
CalculatedControlAscentTimeout := UDINT_TO_TIME(REAL_TO_UDINT(
    LIMIT(CST_TimeoutMinDistance_M, ControlAscentDistance_M, CST_TimeoutMaxDistance_M)
    / CST_MinSpeed_Mps * CST_ControlAscentMargin * CST_SecToMs));

// ⏱️ Integrateurs de temps de montee effective (anti-pompage homme-mort)
IF (ExtractionState = E_ExtractionAssistState.CLOSING_BUCKET) AND MotionRequestActive AND (MotionDirection = 1) THEN
    BucketCloseTimerAcc := BucketCloseTimerAcc + CycleTime;
    IF BucketCloseTimerAcc >= CfgBucketCloseTimeout THEN
        TimeoutBucketCloseFault := TRUE;
    END_IF;
END_IF;

IF (ExtractionState = E_ExtractionAssistState.CONTROL_ASCENT) AND MotionRequestActive AND (MotionDirection = 1) THEN
    ControlAscentTimerAcc := ControlAscentTimerAcc + CycleTime;
    IF ControlAscentTimerAcc >= CalculatedControlAscentTimeout THEN
        TimeoutControlAscentFault := TRUE;
    END_IF;
END_IF;

// Etat physique des causes treuil/benne : conditionne l'acquittement des latches a cause persistante (F2).
CausesPhysiquesEffacees := NOT BucketError AND NOT WinchSyncError
                        AND PositionsValid AND M1MeasuredSpeedValid AND M2MeasuredSpeedValid;
IF ResetEdge.Q AND NOT ErrorCausePresent AND NOT MotionRequestActive THEN
    // Latches sans cause physique persistante (timeouts, backstop) : acquittables sur simple front Reset.
    TimeoutBucketCloseFault   := FALSE;
    TimeoutControlAscentFault := FALSE;
    BucketCloseTimerAcc       := T#0ms;
    ControlAscentTimerAcc     := T#0ms;
    StepAtFaultCaptured       := FALSE;
    ExtractionState := E_ExtractionAssistState.WAIT_BOTTOM_CONFIRMATION;
    // Latches de cause physique : acquittables SEULEMENT si l'entree de defaut est revenue saine (F2).
    IF CausesPhysiquesEffacees THEN
        BucketErrorFault      := FALSE;
        SyncOrSpeedErrorFault := FALSE;
    END_IF;
END_IF;

instCauses[1].Active   := BucketErrorFault;
instCauses[1].Latching := TRUE;
instCauses[1].Texte    := 'Defaut sous-systeme benne pendant fermeture';

instCauses[2].Active   := SyncOrSpeedErrorFault;
instCauses[2].Latching := TRUE;
instCauses[2].Texte    := 'Defaut synchro ou capteurs treuils pendant remontee';

instCauses[3].Active   := ErrorCausePresent;
instCauses[3].Latching := TRUE;
instCauses[3].Texte    := 'Parametrage distance de controle ou backstop invalide';

instCauses[4].Active   := TimeoutBucketCloseFault;
instCauses[4].Latching := TRUE;
instCauses[4].Texte    := 'Depassement backstop fermeture benne';

instCauses[5].Active   := TimeoutControlAscentFault;
instCauses[5].Latching := TRUE;
instCauses[5].Texte    := 'Depassement tempo decollage controle';

// Appel du socle de défaut
instFault(Enable := Enable, Reset := Reset, Causes := instCauses);
Fault := instFault.Fault;

// 📸 Capture ordonnee de StepAtFault (D2). Les defauts leves dans le CASE se figent au site du
// latch (voir §3) ; ce bloc ne couvre que les defauts detectes en §1 (backstop, timeout, parametrage),
// ou ExtractionState/PrevState sont encore l'etape reelle. StepAtFaultCaptured evite l'ecrasement.
ErrorEdge(CLK := Fault.Error);
IF ErrorEdge.Q AND NOT StepAtFaultCaptured THEN
    StepAtFault := PrevState;
    StepAtFaultCaptured := TRUE;
ELSIF ResetEdge.Q AND NOT ErrorCausePresent AND NOT MotionRequestActive THEN
    StepAtFault := E_ExtractionAssistState.WAIT_BOTTOM_CONFIRMATION;
END_IF;
{endregion}

{region "§2 Gate neutralisation"}
// 🛑 2. GATE
IF NOT Enable OR NOT PowerContactorEngaged THEN
    Ready := FALSE;
    Lifecycle.Busy := FALSE;
    Lifecycle.Done := FALSE;
    BucketCloseRequest := FALSE;
    AscentPermit := FALSE;
    ExtractionControlActive := FALSE;
    BottomConfirmationConsumed := FALSE;
    ExtractionState := E_ExtractionAssistState.WAIT_BOTTOM_CONFIRMATION;
    // StepAtFault / StepAtFaultCaptured NON reinitialises ici : l'etape figee au defaut reste
    // lisible pour l'IHM/diagnostic apres un cycle Enable OFF->ON ; seul un front Reset l'efface.
    PrevState := E_ExtractionAssistState.WAIT_BOTTOM_CONFIRMATION;
    BucketCloseTimerAcc := T#0ms;
    ControlAscentTimerAcc := T#0ms;
    OperatorActionId := 0;
    OperatorAction := '';
    RETURN;
END_IF;

Ready := Enable AND NOT Fault.Latched;
{endregion}

{region "§3 Machine etat fermeture remontee"}
BucketCloseRequest := FALSE;
AscentPermit := FALSE;
ExtractionControlActive := FALSE;
BottomConfirmationConsumed := FALSE;
Lifecycle.Busy := FALSE;
Lifecycle.Done := FALSE;

// Ascending assistee reellement demandee : sens ascending + mode maintenance (H5, double garde vs Enable PRG_03).
AssistPermit := MotionRequestActive AND (MotionDirection = 1)
            AND (Mode = E_Mode.MAINT_N1 OR Mode = E_Mode.MAINT_N2);
// Entrees [SAFE] saines : coupure meme-scan des permis si defaut treuil/synchro (H2), avant meme le latch.
AscentControlSafe := NOT WinchSyncError AND PositionsValid AND M1MeasuredSpeedValid AND M2MeasuredSpeedValid;
AscentNominalSafe := NOT WinchSyncError AND PositionsValid;

// Garde-fou non-redemarrage auto : un defaut latche non acquitte verrouille la machine
// d'etat en ERROR_HOLD, meme si la vue live Fault.Error retombe (cause disparue).
IF Fault.Error OR Fault.Latched THEN
    ExtractionState := E_ExtractionAssistState.ERROR_HOLD;
    OperatorActionId := 16#0280;
    OperatorAction := 'Vérifier la benne et les treuils puis réarmer avant de reprendre.';
ELSE
    CASE ExtractionState OF
        E_ExtractionAssistState.WAIT_BOTTOM_CONFIRMATION:
            IF BottomPositionConfirmed THEN
                ExtractionState := E_ExtractionAssistState.READY_TO_CLOSE;
            ELSE
                OperatorActionId := 16#0200;
                OperatorAction := 'Confirmer que la benne est posée au fond avant extraction.';
            END_IF;

        E_ExtractionAssistState.READY_TO_CLOSE:
            Ready := TRUE;
            OperatorActionId := 16#0201;
            OperatorAction := 'Demander la montée pour fermer la benne.';
            IF MotionRequestActive AND (MotionDirection = 1) THEN
                BottomConfirmationConsumed := TRUE;
                BucketCloseTimerAcc := T#0ms;   // ⏱️ RAZ a l'entree exacte de CLOSING_BUCKET
                ExtractionState := E_ExtractionAssistState.CLOSING_BUCKET;
            END_IF;

        E_ExtractionAssistState.CLOSING_BUCKET:
            Lifecycle.Busy := TRUE;
            BucketCloseRequest := AssistPermit AND NOT BucketError; // coupure meme-scan sur defaut benne (H2)
            // Autorisation de montee pendant la fermeture : la benne se ferme en montant.
            // Consommee par l'arbitrage (PRG_04) comme permis de montee assistee (H2).
            AscentPermit := AssistPermit AND AscentControlSafe;
            OperatorActionId := 16#0202;
            OperatorAction := 'Maintenir la montée : fermeture de la benne en cours.';
            IF BucketError THEN
                IF NOT StepAtFaultCaptured THEN
                    StepAtFault := ExtractionState;
                    StepAtFaultCaptured := TRUE;
                END_IF;
                BucketErrorFault := TRUE;
            ELSIF BucketIsClosed AND NOT BucketBusy THEN
                ControlStartM1Position_M := M1Position_M;
                ControlStartM2Position_M := M2Position_M;
                ControlAscentTimerAcc := T#0ms;   // ⏱️ RAZ a l'entree exacte de CONTROL_ASCENT
                ExtractionState := E_ExtractionAssistState.CONTROL_ASCENT;
            END_IF;

        E_ExtractionAssistState.CONTROL_ASCENT:
            Lifecycle.Busy := TRUE;
            AscentPermit := AssistPermit AND AscentControlSafe; // coupure meme-scan sur defaut synchro/capteurs (H2)
            ExtractionControlActive := AscentPermit;            // plafond palier 1 suit le permis de montee
            OperatorActionId := 16#0203;
            OperatorAction := 'Maintenir la montée : contrôle charge au palier minimal.';
            IF NOT AscentControlSafe THEN
                IF NOT StepAtFaultCaptured THEN
                    StepAtFault := ExtractionState;
                    StepAtFaultCaptured := TRUE;
                END_IF;
                SyncOrSpeedErrorFault := TRUE;
            ELSIF (M1Position_M >= (ControlStartM1Position_M + ControlAscentDistance_M))
               AND (M2Position_M >= (ControlStartM2Position_M + ControlAscentDistance_M)) THEN
                ExtractionState := E_ExtractionAssistState.NOMINAL_ASCENT;
            END_IF;

        E_ExtractionAssistState.NOMINAL_ASCENT:
            Lifecycle.Busy := TRUE;
            AscentPermit := AssistPermit AND AscentNominalSafe; // coupure meme-scan sur defaut synchro/position (H2)
            OperatorActionId := 16#0204;
            OperatorAction := 'Maintenir la montée : extraction en cours.';
            IF NOT AscentNominalSafe THEN
                IF NOT StepAtFaultCaptured THEN
                    StepAtFault := ExtractionState;
                    StepAtFaultCaptured := TRUE;
                END_IF;
                SyncOrSpeedErrorFault := TRUE;
            END_IF;

        E_ExtractionAssistState.ERROR_HOLD:
            ;
    END_CASE;
END_IF;

// 💾 Memorisation de la phase precedente en toute fin de scan (capture StepAtFault fiable)
PrevState := ExtractionState;
{endregion}

END_FUNCTION_BLOCK
